        IF (CartesianVx > VXThreshold)
           AND (CartesianForcefX > FXThreshold) THEN

            CASE stFromUnity.nGameStatus OF

                0: // Not playing
                    stJointTargetTorque.M1 := 0.0;

                1: // Light bin
                    stJointTargetTorque.M1 := 0.0;

                2: // Medium bin
                    stJointTargetTorque.M1 := 7.0;

                3: // Heavy bin
                    stJointTargetTorque.M1 := 15.0;

                ELSE
                    stJointTargetTorque.M1 := 0.0;

            END_CASE;


        (****************************************************
            CONDITION 2: NEGATIVE X MOVEMENT

            Both Vx and Fx must be negative
            and below their negative thresholds.

            Apply POSITIVE resistance.
        *****************************************************)

        ELSIF (CartesianVx < -VXThreshold)
              AND (CartesianForcefX < -FXThreshold) THEN

            CASE stFromUnity.nGameStatus OF

                0: // Not playing
                    stJointTargetTorque.M1 := 0.0;

                1: // Light bin
                    stJointTargetTorque.M1 := 0.0;

                2: // Medium bin
                    stJointTargetTorque.M1 := -7.0;

                3: // Heavy bin
                    stJointTargetTorque.M1 := -15.0;

                ELSE
                    stJointTargetTorque.M1 := 0.0;

            END_CASE;

        ELSE

            // Force and velocity conditions not satisfied
            stJointTargetTorque.M1 := 0.0;

        END_IF;
	
	ELSE
		
		GVL_HMI.bLaunchGameSorter:= FALSE;
	
	END_IF

  

END_IF;

END_FUNCTION_BLOCK

// ---- POUs/Crazy Car/FB_CrazyCarGame.TcPOU
FUNCTION_BLOCK FB_CrazyCarGame

VAR_INPUT
    bEnable                   : BOOL;
    stCartesianPosePercentage : ST_CartesianPose;
    fWristAngleDeg            : LREAL;
    CartesianVtheta           : LREAL;
    CartesianMtheta           : LREAL;
END_VAR

VAR_OUTPUT
    stJointTargetTorque : ST_JointTorque;
END_VAR

VAR
    // =====================================================
    // UNITY COMMUNICATION
    // =====================================================

    stToUnity   : ST_CrazyCarToUnity;
    stFromUnity : ST_UnityToCrazyCar;


    // =====================================================
    // RESISTANCE LEVELS
    // =====================================================

    TorqueTaxi  : LREAL := 0.0;
    TorqueVan   : LREAL := 20.0;
    TorqueTruck : LREAL := 40.0;

    TorqueSign  : LREAL := 1.0;

    fTorque : LREAL := 0.0;


    // =====================================================
    // VELOCITY FILTER
    // =====================================================

    fVthetaFiltered : LREAL := 0.0;

    fFilterTime : LREAL := 0.015;

    fTaskCycleTime : LREAL := 0.01;


    // =====================================================
    // VELOCITY DEAD ZONE AND TRANSITION
    //
    // Assumes CartesianVtheta is in deg/s
    // =====================================================

    fVelocityDeadband : LREAL := 10.0;

    fVelocityFull : LREAL := 30.0;


    // =====================================================
    // SMOOTH RESISTANCE
    // =====================================================

    fVelocityMagnitude : LREAL := 0.0;

    fVelocityFactor : LREAL := 0.0;

    fSmoothFactor : LREAL := 0.0;

    fTorqueTarget : LREAL := 0.0;

    fTorqueCommand : LREAL := 0.0;


    // =====================================================
    // APPLICATION TORQUE SLEW LIMIT
    //
    // Units must match the game torque command per second.
    // =====================================================

    fTorqueRateLimit : LREAL := 100.0;

    fMaxTorqueStep : LREAL := 0.0;

    fTorqueDifference : LREAL := 0.0;


    // =====================================================
    // INITIAL BENCH-TEST LIMITS
    //
    // Keep motor output disabled while validating the logic.
    // fMaxGameTorque is an experimental command bound,
    // NOT a validated safe human-interaction torque.
    // =====================================================

    bEnableResistanceOutput : BOOL := FALSE;

    fMaxGameTorque : LREAL :=40.0;

END_VAR

(************************************************************
    CRAZY CAR GAME - CONTINUOUS SMOOTH RESISTANCE

    Unity status:
        0 = Menu / Popup
        1 = Taxi
        2 = Van
        3 = Truck

    Objectives:
        1. Zero resistance near stationary velocity
        2. Smooth resistance transition
        3. Approximately constant resistance during motion
        4. Avoid binary torque switching
        5. Limit the commanded torque rate
*************************************************************)


// ==========================================================
// 1. DEFAULT OUTPUTS
// ==========================================================

stJointTargetTorque.M1 := 0.0;
stJointTargetTorque.M2 := 0.0;
stJointTargetTorque.M3 := 0.0;

stToUnity.GameIsActive := FALSE;

fTorque := 0.0;
fTorqueTarget := 0.0;


// ==========================================================
// 2. CHECK GAME ENABLE
// ==========================================================

IF bEnable AND NOT stFromUnity.bGameClosed THEN

    // Send data to Unity

    stToUnity.fY :=
        LREAL_TO_REAL(stCartesianPosePercentage.Y);

    stToUnity.fWristAngle :=
        LREAL_TO_REAL(fWristAngleDeg);

    stToUnity.GameIsActive := TRUE;


    // ======================================================
    // 3. READ VEHICLE RESISTANCE
    // ======================================================

    CASE stFromUnity.nGameStatus OF

        1:
            fTorque := TorqueTaxi;

        2:
            fTorque := TorqueVan;

        3:
            fTorque := TorqueTruck;

        ELSE
            fTorque := 0.0;

    END_CASE;


    // ======================================================
    // 4. FILTER WRIST VELOCITY
    // ======================================================

    IF (fTaskCycleTime > 0.0)
       AND (fFilterTime >= 0.0) THEN

        fVthetaFiltered :=
            fVthetaFiltered
            +
            (
                fTaskCycleTime /
                (fFilterTime + fTaskCycleTime)
            )
            *
            (CartesianVtheta - fVthetaFiltered);

    ELSE

        fVthetaFiltered := 0.0;

    END_IF;


    // ======================================================
    // 5. CALCULATE VELOCITY MAGNITUDE
    // ======================================================

    fVelocityMagnitude := ABS(fVthetaFiltered);


    // ======================================================
    // 6. CALCULATE CONTINUOUS VELOCITY FACTOR
    //
    // Dead zone:          Factor = 0
    // Transition region:  Factor = 0..1
    // Full movement:      Factor = 1
    // ======================================================

    fVelocityFactor := 0.0;

    IF fVelocityFull > fVelocityDeadband THEN

        IF fVelocityMagnitude <= fVelocityDeadband THEN

            fVelocityFactor := 0.0;

        ELSIF fVelocityMagnitude >= fVelocityFull THEN

            fVelocityFactor := 1.0;

        ELSE

            fVelocityFactor :=
                (fVelocityMagnitude - fVelocityDeadband)
                /
                (fVelocityFull - fVelocityDeadband);

        END_IF;

    END_IF;


    // ======================================================
    // 7. SMOOTHSTEP FUNCTION
    //
    // Smooth transition from 0 to 1.
    //
    // f(x) = 3*x*x - 2*x*x*x
    //
    // This avoids an abrupt slope change at the
    // beginning and end of the transition region.
    // ======================================================

    fSmoothFactor :=
        fVelocityFactor
        *
        fVelocityFactor
        *
        (3.0 - 2.0 * fVelocityFactor);


    // ======================================================
    // 8. CALCULATE TARGET RESISTANCE
    //
    // Preserve your existing motor sign convention.
    // Verify that the physical wrist torque opposes motion.
    // ======================================================

    IF fVthetaFiltered > fVelocityDeadband THEN

        fTorqueTarget :=
            TorqueSign
            *
            fTorque
            *
            fSmoothFactor;

    ELSIF fVthetaFiltered < -fVelocityDeadband THEN

        fTorqueTarget :=
            -TorqueSign
            *
            fTorque
            *
            fSmoothFactor;

    ELSE

        fTorqueTarget := 0.0;

    END_IF;


    // ======================================================
    // 9. LIMIT GAME TORQUE MAGNITUDE
    //
    // Experimental bench-test limit.
    // ======================================================

    IF bEnableResistanceOutput
       AND (fMaxGameTorque > 0.0) THEN

        fTorqueTarget :=
            MAX(
                -fMaxGameTorque,
                MIN(fMaxGameTorque, fTorqueTarget)
            );

    ELSE

        fTorqueTarget := 0.0;

    END_IF;


    // ======================================================
    // 10. APPLICATION-LEVEL TORQUE SLEW LIMIT
    //
    // Prevent large command changes within one PLC cycle.
    // ======================================================

    fMaxTorqueStep :=
        MAX(0.0, fTorqueRateLimit)
        *
        MAX(0.0, fTaskCycleTime);

    fTorqueDifference :=
        fTorqueTarget - fTorqueCommand;


    IF fTorqueDifference > fMaxTorqueStep THEN

        fTorqueCommand :=
            fTorqueCommand + fMaxTorqueStep;

    ELSIF fTorqueDifference < -fMaxTorqueStep THEN

        fTorqueCommand :=
            fTorqueCommand - fMaxTorqueStep;

    ELSE

        fTorqueCommand := fTorqueTarget;

    END_IF;


    // ======================================================
    // 11. TRANSFER TORQUE TO WRIST MOTORS
    // ======================================================

    IF bEnableResistanceOutput THEN

        stJointTargetTorque.M2 := fTorqueCommand;
        stJointTargetTorque.M3 := fTorqueCommand;

    ELSE

        stJointTargetTorque.M2 := 0.0;
        stJointTargetTorque.M3 := 0.0;

        fTorqueCommand := 0.0;

    END_IF;


ELSE

    // ======================================================
    // 12. GAME DISABLED OR CLOSED
    // ======================================================

    IF bEnable AND stFromUnity.bGameClosed THEN

        GVL_HMI.bLaunchGameCrazyCar := FALSE;

    END_IF;


    stToUnity.GameIsActive := FALSE;

    fTorque := 0.0;
    fTorqueTarget := 0.0;
    fTorqueCommand := 0.0;

    fVthetaFiltered := 0.0;

    fVelocityMagnitude := 0.0;
    fVelocityFactor := 0.0;
    fSmoothFactor := 0.0;

    fTorqueDifference := 0.0;

END_IF;

END_FUNCTION_BLOCK

// ---- POUs/Firrfly Game/FB_FireflyGame.TcPOU
FUNCTION_BLOCK FB_FireflyGame
VAR_INPUT
    bEnable                   : BOOL;
    stCartesianPosePercentage : ST_CartesianPose; // from Kinematics: X -100..+100 %, Y 0..100 % (0..370 mm)
END_VAR
VAR_OUTPUT
    stJointTargetTorque : ST_JointTorque;  // always 0: Firefly is motion-only, no actuation
    nGameStatus         : INT;             // Unity game status, for MAIN / HMI
    bExitRequested      : BOOL;            // TRUE for ONE PLC cycle when Exit is pressed in Unity
    bWrongFlowerEvent   : BOOL;            // TRUE for ONE PLC cycle per wrong flower (for later haptics)
END_VAR
VAR
    stToUnity   : ST_FireflyToUnity;
    stFromUnity : ST_FireflyFromUnity;

    // Calibration: robot percent (from Kinematics) at home, and travel either side of home
    // that brings the firefly to the edge of the garden (= +/-100 % in Unity).
    fXHome      : REAL := 0.0;    // X percent at home (middle of the workspace)
    fYHome      : REAL := 50.0;   // Y percent at home (middle of 0..370 mm = 185 mm)
    fXHalfRange : REAL := 50.0;   // X: lower this if X needs less motion than Y
    fYHalfRange : REAL := 25.0;   // Y: +/-25 % = 50 % of the Y range of motion in total

    rtExit  : R_TRIG;
    rtWrong : R_TRIG;
    fXRaw   : REAL;
    fYRaw   : REAL;
END_VAR

// Firefly is motion-only: never apply torque.
stJointTargetTorque.M1 := 0.0;
stJointTargetTorque.M2 := 0.0;
stJointTargetTorque.M3 := 0.0;

IF bEnable THEN
    fXRaw := TO_REAL(stCartesianPosePercentage.X);
    fYRaw := TO_REAL(stCartesianPosePercentage.Y);
    // Home -> 0 %, home +/- half range -> +/-100 %, clamped so the firefly stays inside the garden.
    stToUnity.fX := LIMIT(-100.0, (fXRaw - fXHome) / MAX(fXHalfRange, 0.1) * 100.0, 100.0);
    stToUnity.fY := LIMIT(-100.0, (fYRaw - fYHome) / MAX(fYHalfRange, 0.1) * 100.0, 100.0);
ELSE
    stToUnity.fX := 0.0;   // firefly waits on the home flower
    stToUnity.fY := 0.0;
END_IF

// Unity's pulses -> one-cycle events for MAIN (each new pulse = a new rising edge).
rtExit(CLK := stFromUnity.bExitPressed);
rtWrong(CLK := stFromUnity.bWrongFlower);
bExitRequested    := rtExit.Q;
bWrongFlowerEvent := rtWrong.Q;
nGameStatus       := stFromUnity.nGameStatus;

END_FUNCTION_BLOCK

// ---- POUs/FB_ForceTorqueSensor.TcPOU
FUNCTION_BLOCK FB_ForceTorqueSensor
VAR_IN_OUT
 CartesianState : ST_CartesianState;
 
END_VAR
VAR_INPUT
	CartesianPosAdditionalParameter :ST_CartesianAdditionalParametes;
END_VAR
VAR
    eState : E_CalibrationState :=  E_CalibrationState.INIT;
    tWait  : TON;
	FxTemp : LREAL;
	FyTemp : LREAL;
	MzTemp : LREAL;
	OffsetRawFx: LINT;
	OffsetRawFy: LINT;
	OffsetRawMz: LINT;
	sumFx: LINT;
	sumFy: LINT;
	sumMz: LINT;
	nSample: INT;
	rTrigZero : R_TRIG;
	Theta1: LREAL;
	Theta2: LREAL;
	Theta3: LREAL;
END_VAR
VAR CONSTANT
    CMD_STOP   : DWORD := 16#0000000C;
    CMD_FILTER : DWORD := 16#00050108;  // 1st-order LPF, 100 Hz
    CMD_START  : DWORD := 16#0000000B;
    FORCE_DIV  : REAL := 50.0;     // RFT60-HA01 force divider
	TORQUE_DIV : REAL := 2000.0;   // RFT60-HA01 torque divider
	CostanstAngleBetweenFTSensorAndXdirection : LREAL := 30.0; // Unit Degree
	CostanstAngleBetweenFTSensorAndYdirection : LREAL := 30.0; // Unit Degree
	ZeroingSample : INT := 100;
	
END_VAR



CASE eState OF
E_CalibrationState.INIT:
    GVL_ForceTorqueSensor.ConfigParameter := CMD_STOP;
    tWait(IN := TRUE, PT := T#1000MS);
    IF tWait.Q THEN tWait(IN := FALSE); eState := E_CalibrationState.SET_FILTER; END_IF

E_CalibrationState.SET_FILTER:
   GVL_ForceTorqueSensor.ConfigParameter := CMD_FILTER;
    tWait(IN := TRUE, PT := T#1000MS);
    IF tWait.Q THEN tWait(IN := FALSE); eState := E_CalibrationState.START; END_IF

E_CalibrationState.START:
    GVL_ForceTorqueSensor.ConfigParameter := CMD_START;
    eState := E_CalibrationState.WaitingforCalibrationButton;
	sumFx := 0; sumFy := 0;  sumMz := 0;
	
E_CalibrationState.WaitingforCalibrationButton:

rTrigZero(CLK := GVL_HMI.StartCalibrationButton);

IF rTrigZero.Q THEN

    
   
    GVL_HMI.StartCalibrationButton := FALSE;
	eState := E_CalibrationState.ZEROING;
	sumFx := 0;
	sumFy := 0;
	sumMz := 0;
	nSample := 0;
	tWait(IN := FALSE);   // reset timer

END_IF

	
E_CalibrationState.ZEROING:
   

	tWait(IN := TRUE, PT := T#2000MS);          // let streaming/filter settle first
    IF tWait.Q THEN
        sumFx := sumFx + GVL_ForceTorqueSensor.RawFx;
        sumFy := sumFy + GVL_ForceTorqueSensor.RawFy;
        sumMz := sumMz + GVL_ForceTorqueSensor.RawMz;
        nSample := nSample + 1;
        IF nSample >= ZeroingSample THEN
            OffsetRawFx := sumFx / ZeroingSample;
            OffsetRawFy := sumFy / ZeroingSample;
            OffsetRawMz := sumMz / ZeroingSample;
            eState := E_CalibrationState.RUNNING;
        END_IF
    END_IF



E_CalibrationState.RUNNING:
IF GVL_HMI.StartCalibrationButton THEN
	 GVL_HMI.StartCalibrationButton := FALSE;

    sumFx := 0;
    sumFy := 0;
    sumMz := 0;
    nSample := 0;

    tWait(IN := FALSE);

    eState := E_CalibrationState.ZEROING;
END_IF
// All Angles that is used for rotational frames;
Theta1:= CostanstAngleBetweenFTSensorAndXdirection;   //UNIT: degree   Shift for F/t Sensor, it is related to design and I got from SOLIDWORKS// this number is constant;
Theta2 := -CartesianPosAdditionalParameter.BetaIncremental; // UNIT: degree  the angle between frame x,y with refrence
Theta3 := -Cartesianstate.Position.Theta; //UNIT: degree  the wrist angle between x-frame of wrist with x-frame of reference
//
    FxTemp := LINT_TO_REAL(GVL_ForceTorqueSensor.RawFx- OffsetRawFx) / FORCE_DIV;
    FyTemp := LINT_TO_REAL(GVL_ForceTorqueSensor.RawFy-OffsetRawFy) / FORCE_DIV;
    MzTemp := LINT_TO_REAL(GVL_ForceTorqueSensor.RawMz-OffsetRawMz) / TORQUE_DIV;
	CartesianState.Force.Fx :=-( FxTemp * COS((Theta1 + Theta2 + Theta3)*(PI / 180.0))-
	FyTemp * SIN((Theta1 + Theta2 + Theta3)*(PI / 180.0)));
	
	GVL_HMI.Fx_HMI := CartesianState.Force.Fx ; // Display in HMI
	
	CartesianState.Force.Fy := -(FxTemp * SIN((Theta1 + Theta2 + Theta3)*(PI / 180.0))+
	FyTemp * COS((Theta1 + Theta2 + Theta3)*(PI / 180.0)));
	
	GVL_HMI.Fy_HMI := CartesianState.Force.Fy; // Display in HMI
	CartesianState.Force.Mtheta := MzTemp ;
	GVL_HMI.Mz_HMI := CartesianState.Force.Mtheta*1000;  // Display in HMI //Unit : mNM




END_CASE

IF eState = E_CalibrationState.RUNNING THEN
	GVL_HMI.UserSecuringButton_HMI := TRUE;
	ELSE
	GVL_HMI.UserSecuringButton_HMI := FALSE;	
END_IF

END_FUNCTION_BLOCK

// ---- POUs/HMI_FunBlock/MicroswitchCheck.TcPOU
FUNCTION_BLOCK MicroswitchCheck
VAR_INPUT
END_VAR
VAR_OUTPUT
END_VAR
VAR
	SwTheta1: BOOL;
	SwTheta2: BOOL;
	SwR1: BOOL;
	SwR2: BOOL;
	SwBeta1: BOOL;
	SwBeta2: BOOL;
END_VAR

SwTheta1 	 := (GVL_MicroSwitch.dwMicroSwitchDriverA AND 16#00020000) <> 0;  (* bit 0 *)
SwTheta2     := (GVL_MicroSwitch.dwMicroSwitchDriverA AND 16#00010000) <> 0;  (* bit 1 *)
SwR1    	 := (GVL_MicroSwitch.dwMicroSwitchDriverB AND 16#00080000) <> 0;  (* bit 0 *)
SwR2  		 := (GVL_MicroSwitch.dwMicroSwitchDriverB AND 16#00040000) <> 0;  (* bit 1 *)
SwBeta1      := (GVL_MicroSwitch.dwMicroSwitchDriverB AND 16#00020000) <> 0;  (* bit 2 *)
SwBeta2      := (GVL_MicroSwitch.dwMicroSwitchDriverB AND 16#00010000) <> 0;  (* bit 3 *)

IF SwTheta1 THEN
GVL_HMI.CheckMicroswitchWristLeft := TRUE;
	
END_IF

IF SwTheta2 THEN
GVL_HMI.CheckMicroswitchWristRight := TRUE;
	
END_IF

IF SwR1 THEN
GVL_HMI.CheckMicroswitchLinearMax := TRUE;
	
END_IF

IF SwR2 THEN
GVL_HMI.CheckMicroswitchLinearMin := TRUE;
	
END_IF

IF SwBeta1 THEN
GVL_HMI.CheckMicroswitchRotationRight := TRUE;
	
END_IF

IF SwBeta2 THEN
GVL_HMI.CheckMicroswitchRotationLeft := TRUE;
	
END_IF

IF GVL_HMI.CheckMicroswitchWristLeft AND GVL_HMI.CheckMicroswitchWristRight AND GVL_HMI.CheckMicroswitchLinearMax AND GVL_HMI.CheckMicroswitchLinearMin AND GVL_HMI.CheckMicroswitchRotationRight AND GVL_HMI.CheckMicroswitchRotationLeft THEN
GVL_HMI.ContinueToHoming := TRUE;

END_IF

END_FUNCTION_BLOCK

// ---- POUs/HMI_FunBlock/FB_UserSecuring.TcPOU
FUNCTION_BLOCK FB_UserSecuring
VAR_INPUT
END_VAR
VAR_OUTPUT
END_VAR
VAR
END_VAR

IF GVL_HMI.check1 AND GVL_HMI.check2 AND GVL_HMI.check3 AND GVL_HMI.check4 AND GVL_HMI.check5 AND GVL_HMI.check6 THEN
	
GVL_HMI.ContinueTOWorkspaceLimits := TRUE;
ELSE
	
GVL_HMI.ContinueTOWorkspaceLimits := FALSE;

END_IF

END_FUNCTION_BLOCK

// ---- POUs/FB_TherapyManager.TcPOU
FUNCTION_BLOCK FB_TherapyManager

VAR_INPUT
	Enable         : BOOL;
    Config         : ST_TherapyConfig;       // The struct we just built!
    ActualJoints    : ST_JointState;        // Feedback: Joint q, q_dot, M
    ActualCartesian : ST_CartesianState;    // Feedback: Cartesian Pose, Vel, Force
    TargetCartesian : ST_CartesianTarget;   // Target: Cartesian Pose, Vel, Force setpoints
    SimpleJointTorqueObtainedFromGames : ST_JointTorque;
    fbKinematics    : REFERENCE TO FB_RobotKinematics;
	WallSetPointXandY : ARRAY[1..4, 1..2] OF LREAL;
END_VAR
VAR_OUTPUT
	TargetJointsTorque    : ST_JointTorque;        // Output for CST Mode
	//TargetMode      : En_TargetMode;              // Drive mode (eCSP, eCSV, eCST)
    //  Out_Positions  : ST_JointPositions;      // Output for CSV Mode
END_VAR
VAR
	// 1. The Expert Math Blocks
    fbImpedance    : FB_ImpedanceController;
    fbAdmittance   : FB_AdmittanceController;
	fbForceYield : FB_ForceController;
    fbDynamics     : FB_DynamicsCompensator;
    
    // 2. Internal Routing Variables
    TherapyForces   : ST_CartesianForces;             // Cartesian Space (End-Effector force)
    TherapyTorque   : ST_JointTorque;                 // Joint Space (Therapy motor torque)
    CompTorque      : ST_JointTorque;                 // Joint Space (Hardware compensation torque)
	timerHold : TON;
	
	// Wall Variables
	WallTorque : ST_JointTorque;
	fbVirtualWall : FB_VirtuallWall;
	bWallInContact : BOOL;
	WallCartesianForce: ST_CartesianForces;
	MotionState: INT := 1;
	//cycle: INT;
	CycleMotion: INT :=1;
	
	
	fbMicroswitchCheck : MicroswitchCheck;   // Delete this after cycling test
	fbStopM1 : MC_Stop;
	fbStopM2 : MC_Stop;
	fbStopM3 : MC_Stop;
	firsttime: BOOL := TRUE;
END_VAR
VAR CONSTANT
    // Zero constants for clean single-line memory resets
    cZeroTorque : ST_JointTorque    := (M1 := 0.0, M2 := 0.0, M3 := 0.0);
    cZeroForces : ST_CartesianForces := (Fx := 0.0, Fy := 0.0, Mtheta := 0.0);
END_VAR

// =========================================================
// 1. SAFETY DISABLE GUARD
// =========================================================
IF NOT Enable THEN
    TargetJointsTorque := cZeroTorque;
	
   
    RETURN;
END_IF

// =========================================================
// 2. CLEAR INTERMEDIATE BUFFERS (PREVENT STALE DATA LEAKS)
// =========================================================
TherapyForces := cZeroForces;
TherapyTorque := cZeroTorque;
WallTorque := cZeroTorque;
CompTorque    := cZeroTorque;

// =========================================================
// 3. PRIMARY CONTROLLER ROUTING
// =========================================================
CASE Config.ControllerType OF

    E_ControllerType.ControlNone:
        TherapyTorque := SimpleJointTorqueObtainedFromGames;
		
		(*

    E_ControllerType.ControlImpedance:
        // Step A: Virtual spring-damper computes interaction forces
        fbImpedance(
            Stiffness   := Config.Stiffness_K,
            Damping     := Config.Damping_D,
            ActualPose  := ActualCartesian.Position,
            TargetPose  := TargetCartesian.Position,
            ActualVel   := ActualCartesian.Velocity,
            TargetVel   := TargetCartesian.Velocity,
            OutputForce => TherapyForces
        );
        
        // Step B: Map Cartesian Force -> Joint Torque via J^T
        TherapyTorque := fbKinematics.ApplyJacobianTranspose(Force := TherapyForces);

    E_ControllerType.ControlAdmittance:
        // Measured patient forces generate target positions / velocities
        fbAdmittance(
            TherapyMode     := Config.TherapyMode,
            VirtualMass     := Config.Mass_M,
            VirtualDamp     := Config.Damping_D,
            MeasuredForces  := ActualCartesian.Forces,
            TargetForces    := TargetCartesian.Forces,
            ActualPose      := ActualCartesian.Position,
            TargetPosition  => TargetJoints.Position
        );

    E_ControllerType.ControlForce:
        // Generic Yield-Threshold / Breakaway Force Controller
        fbForceYield(
            ForceThreshold := Config.ForceConfig.Threshold, // Generic resistance force
            VirtualDamping := Config.ForceConfig.Damping,   // Generic motion viscosity
            ActualForce    := ActualCartesian.Forces,
            ActualJoints   := ActualJoints,
            OutputTorque   => TherapyTorque
        );
		*)

END_CASE

// =========================================================
// 4. HARDWARE DYNAMICS COMPENSATION (Joint Space)
// =========================================================

(*

IF Config.FeatureFrictionComp OR Config.FeatureInertiaComp OR Config.FeatureGravityComp THEN
    fbDynamics(
        JointPosition  := ActualJoints.Position,
        JointVelocity  := ActualJoints.Velocity,
        EnableGravity  := Config.FeatureGravityComp,
        EnableFriction := Config.FeatureFrictionComp,
        EnableInertia  := Config.FeatureInertiaComp,
        CompTorque     => CompTorque
    );
END_IF
*)
// Cycle Test
(* 

IF  firsttime THEN
GVL_hmi.CheckMicroswitchLinearMax := FALSE;
GVL_hmi.CheckMicroswitchLinearMin := FALSE;
GVL_hmi.CheckMicroswitchRotationLeft := FALSE;
GVL_hmi.CheckMicroswitchRotationRight := FALSE;
GVL_HMI.CheckMicroswitchWristLeft := FALSE;
GVL_HMI.CheckMicroswitchWristRight := FALSE;
firsttime := FALSE;
END_IF
// Tests
fbMicroswitchCheck();
IF GVL_hmi.CheckMicroswitchLinearMax OR GVL_hmi.CheckMicroswitchLinearMin OR
 GVL_hmi.CheckMicroswitchRotationLeft OR GVL_hmi.CheckMicroswitchRotationRight OR 
 GVL_HMI.CheckMicroswitchWristLeft OR GVL_HMI.CheckMicroswitchWristRight

THEN
 
	fbStopM1(
        Axis      := GVL_Axes.Axis1,
        Execute   := TRUE);   

    fbStopM2(
        Axis      := GVL_Axes.Axis2,
        Execute   := TRUE);

    fbStopM3(
        Axis      := GVL_Axes.Axis3,
        Execute   := TRUE);
END_IF

CASE MotionState OF
	1: // Motor1 +_
		TherapyTorque.M1 := -8.0;
		TherapyTorque.M2 := 0.0;
		TherapyTorque.M3 := 0.0;
		IF ActualCartesian.Position.X> 200.0 THEN
			
		TherapyTorque.M1 :=  0.05* ActualCartesian.Velocity.Vx;
		TherapyTorque.M2 := 0.0;
		TherapyTorque.M3 := 0.0;
		timerHold(IN := TRUE, PT := T#1S);
		
		IF timerHold.Q THEN
            timerHold(IN := FALSE); // Reset the timer so it can be reused later
            MotionState := 2;
        END_IF
			
		END_IF
	2: // linear +
		TherapyTorque.M1 := 0.0;
		TherapyTorque.M2 := 8.0;
		TherapyTorque.M3 := -8.0;
		
		IF ActualCartesian.Position.Y> 300.0 THEN
		TherapyTorque.M1 := 0.0;
		TherapyTorque.M2 :=  - 0.05* ActualCartesian.Velocity.Vy;
		TherapyTorque.M3 :=  0.05* ActualCartesian.Velocity.Vy;
		timerHold(IN := TRUE, PT := T#1S);
		
		IF timerHold.Q THEN
            timerHold(IN := FALSE); // Reset the timer so it can be reused later
            MotionState := 3;
		END_IF
		END_IF
	 3: // Motor1 -
		TherapyTorque.M1 := 8.0;
		TherapyTorque.M2 := 0.0;
		TherapyTorque.M3 := 0.0;
		
		IF ActualCartesian.Position.X< -50.0 THEN
		TherapyTorque.M1 := 0.05* ActualCartesian.Velocity.Vx;
		TherapyTorque.M2:= 0.0;
		TherapyTorque.M3 := 0.0;
		timerHold(IN := TRUE, PT := T#1S);
		
		IF timerHold.Q THEN
            timerHold(IN := FALSE); // Reset the timer so it can be reused later
            MotionState := 4;
		END_IF
		END_IF
	 4: // linear -
		TherapyTorque.M1 := 0.0;
		TherapyTorque.M2 := -8.0;
		TherapyTorque.M3 := 8.0;
		
		
		IF ActualCartesian.Position.Y< 150.0 THEN
		TherapyTorque.M1 := 0.0;
		TherapyTorque.M2 :=  - 0.05* ActualCartesian.Velocity.Vy;
		TherapyTorque.M3 :=  0.05* ActualCartesian.Velocity.Vy;
		timerHold(IN := TRUE, PT := T#1S);
		
		IF timerHold.Q THEN
            timerHold(IN := FALSE); // Reset the timer so it can be reused later
			CycleMotion := CycleMotion+1;
		IF CycleMotion = 500 THEN
            MotionState := 5;
		ELSE
	MotionState := 1;
			
		END_IF
		END_IF
		END_IF
		
		
	 5: 
		TherapyTorque.M1 := 0.0;
		TherapyTorque.M2 := 0.0;
		TherapyTorque.M3 := 0.0;
		
	 
	 
	
END_CASE

*)// Cycle Test

// VirtualWallTorque

fbVirtualWall(
    bEnable     := GVL_HMI.EableVirtuallWall_Planar,
	Endeffectorstatus := ActualCartesian,
	WallSetPointXandY := WallSetPointXandY,
	WallCartesianForce => WallCartesianForce,
	bInContact  => bWallInContact
    
);

WallTorque :=
    fbKinematics.CartesianForceToTorque(
        Force := WallCartesianForce
    );





// =========================================================
// 5. FINAL TORQUE SUMMATION & GLOBAL SAFETY CLAMP
// =========================================================
IF bWallInContact THEN

    // Virtual wall is active:
    // use wall torque only
    TargetJointsTorque.M1 := LIMIT(
        -Config.GlobalForceLimit,
        WallTorque.M1,
        Config.GlobalForceLimit
    );

    TargetJointsTorque.M2 := LIMIT(
        -Config.GlobalForceLimit,
        WallTorque.M2,
        Config.GlobalForceLimit
    );

    TargetJointsTorque.M3 := LIMIT(
        -Config.GlobalForceLimit,
        WallTorque.M3,
        Config.GlobalForceLimit
    );

ELSE

    // No wall contact:
    // normal robot torque
    TargetJointsTorque.M1 := LIMIT(
        -Config.GlobalForceLimit,
        TherapyTorque.M1 + CompTorque.M1,
        Config.GlobalForceLimit
    );

    TargetJointsTorque.M2 := LIMIT(
        -Config.GlobalForceLimit,
        TherapyTorque.M2 + CompTorque.M2,
        Config.GlobalForceLimit
    );

    TargetJointsTorque.M3 := LIMIT(
        -Config.GlobalForceLimit,
        TherapyTorque.M3 + CompTorque.M3,
        Config.GlobalForceLimit
    );

END_IF;

END_FUNCTION_BLOCK

// ---- POUs/FB_ImpedanceController.TcPOU
FUNCTION_BLOCK FB_ImpedanceController
VAR_INPUT
 TherapyMode : E_RehabMode;
 Stiffness   : LREAL;              // Virtual spring K
 Damping     : LREAL;              // Virtual friction D
  
END_VAR



VAR_OUTPUT
    bBusy         : BOOL;
    bError        : BOOL;
    bDone         : BOOL;
//	TherapyTorques : ST_JointTorques;
END_VAR

VAR
	 
    stPointA      : ARRAY [1..3] OF LREAL  ; 
    stPointB      : ARRAY [1..3] OF LREAL  ;
    stPointC      : ARRAY [1..3] OF LREAL  ;
	
    // --- Feedback from Robot (Inputs) ---
    ActX          : LREAL; 
    ActY          : LREAL; 
    ActTheta      : LREAL;
	ActR          : LREAL; // mm
	ActBeta		  : LREAL;
    


    // --- State Machine Logic ---
    iState           : INT := 0;      // Main Step Counter
    iCurrentSegment  : INT := 0;      // 5=Approach, 10=A->B, 20=B->C, 30=C->A
    bAtPointA        : BOOL := FALSE;
    bSegmentDone     : BOOL;
    bWaitEnable      : BOOL;
    
    // --- Timers & Sub-FBs ---
    fbWaitTimer      : TON;           // Timer for resting at corners
    fbKinematic      : FB_RobotKinematics;  // Internal instance to update kinematics
    
    // --- Motion Profile Variables (Trapezoid Generator) ---
    lrS_T            : LREAL;         // Current Distance along path (0 to L)
    lrS_dot          : LREAL;         // Current Velocity (Speed of the "Rabbit")
    lrL_Target       : LREAL;         // Total Length of the current segment

    // --- Geometric Calculations (Approach Phase) ---
    lrApproachStartX : LREAL;
    lrApproachStartY : LREAL;
    lrApproachStartTheta : LREAL;
    lrDX_App, lrDY_App, lrDTh_App, lrL_App : LREAL;

    // --- Geometric Calculations (Triangle Phase) ---
    // Line 1 (A->B)
    lrDX1, lrDY1, lrDTh1, lrL1 : LREAL;
    // Line 2 (B->C)
    lrDX2, lrDY2, lrDTh2, lrL2 : LREAL;
    // Line 3 (C->A)
    lrDX3, lrDY3, lrDTh3, lrL3 : LREAL;

    // --- Impedance Control Targets ---
    SetAppX             : LREAL; // The "Virtual Rabbit" X position
    SetAppY             : LREAL; // The "Virtual Rabbit" Y position
    SetAppTheta         : LREAL; // The "Virtual Rabbit" Theta position
    
    // --- Calculation Results ---
    CalcForces       : ARRAY [1..3] OF LREAL; // [Fx, Fy, Mz] calculated by Impedance
    CalcTorques      : ARRAY [1..3] OF LREAL; // [Tau1, Tau2, Tau3] calculated by Jacobian

    // --- TwinCAT Motion Control Blocks ---
    // Note: I renamed these to 'fbTorqueAxis1' to match the method code we wrote previously
    fbTorqueAxis1    : MC_TorqueControl;
    fbTorqueAxis2    : MC_TorqueControl;
    fbTorqueAxis3    : MC_TorqueControl;

    // --- Safety Parameters ---
    MaxSpeedLimit    : LREAL := 70.0; // Safety velocity limit (mm/s)
    MaxTorqueLimit   : LREAL := 50.0;  // Safety torque limit (Nm)
	
	// 
	lrVmax: LREAL := 10.0; // mm/s
	lrAcc : LREAL := 100.0 ;// mm/ s^2
	
	SetVelAppX      : LREAL;
    SetVelAppY      : LREAL;
    SetVelAppTheta  : LREAL;
	
	// INTERNAL setpoints calculated each cycle
    stCurrentSet  : ARRAY[1..3] OF LREAL; // Target [X, Y, Theta]
	 lrVx_FF, lrVy_FF, lrVTh_FF : LREAL;
	  Ex, Ey, ETheta    : LREAL; // Position Errors
	  lrTorqueSetpoint_Pct : ARRAY[1..3] OF LREAL;
END_VAR

(* This Function block can be used for difference rehabilitation mode
 1- passive motion: actuators create No torque and patient can move the robot
 2- Passive motion + Compensation(solving dynamic of robot)
 3- Resistive or Assistive force
*)

stPointA := GVL_TargetPoints.Target_A;
stPointB := GVL_TargetPoints.Target_B;
stPointC := GVL_TargetPoints.Target_C;


// =========================================================
// 1. KINEMATICS UPDATE (Always Run First)
// =========================================================
// We need ActX/ActY to calculate the spring force error
(*  JUST FOR TEST ELIMINATED
fbKinematic(
	
    q1 := GVL_RobotData.Q1_Actual, 
    q2 := GVL_RobotData.Q2_Actual, 
    q3 := GVL_RobotData.Q3_Actual, 
    X_Dir => ActX, 
    Y_Dir => ActY, 
    Theta => ActTheta,
    R_Dir => ActR,
	Beta => ActBeta    
);
*)

// 

// Update Timer
fbWaitTimer(IN := bWaitEnable, PT := T#120S);

// =========================================================
// 2. STATE MACHINE
// =========================================================
CASE iState OF

    // -----------------------------------------------------
    // STATE 0: INITIALIZATION (Math Setup)
    // -----------------------------------------------------
    0: 
        // 1. Capture Start Position for Approach
        lrApproachStartX     := ActX;
        lrApproachStartY     := ActY;
        lrApproachStartTheta := ActTheta;

        // 2. Calculate Distance to Point A (Approach Vector)
        lrDX_App  := stPointA[1] - lrApproachStartX;
        lrDY_App  := stPointA[2] - lrApproachStartY;
        lrDTh_App := stPointA[3] - lrApproachStartTheta;
        lrL_App   := MAX(0.001, SQRT(lrDX_App*lrDX_App + lrDY_App*lrDY_App));

        // 3. Calculate Triangle Vectors (A->B, B->C, C->A)
        // --- Line 1: A to B ---
        lrDX1  := stPointB[1] - stPointA[1];
        lrDY1  := stPointB[2] - stPointA[2];
        lrDTh1 := stPointB[3] - stPointA[3];
        lrL1   := MAX(0.001, SQRT(lrDX1*lrDX1 + lrDY1*lrDY1));
        
        // --- Line 2: B to C ---
        lrDX2  := stPointC[1] - stPointB[1];
        lrDY2  := stPointC[2] - stPointB[2];
        lrDTh2 := stPointC[3] - stPointB[3];
        lrL2   := MAX(0.001, SQRT(lrDX2*lrDX2 + lrDY2*lrDY2));
        
        // --- Line 3: C to A ---
        lrDX3  := stPointA[1] - stPointC[1];
        lrDY3  := stPointA[2] - stPointC[2];
        lrDTh3 := stPointA[3] - stPointC[3];
        lrL3   := MAX(0.001, SQRT(lrDX3*lrDX3 + lrDY3*lrDY3));

        // Reset Motion
        lrS_T   := 0;
        lrS_dot := 0;
        
        iCurrentSegment := 5; // Start with Approach
        GVL_MessageStaus.MessageStaus := 'Assistive: Guiding to Start Point A.';
        iState  := 5;


    // -----------------------------------------------------
    // STATE 5: APPROACH (Guiding Patient to Point A)
    // -----------------------------------------------------
    5:
        // A. Move the "Virtual Rabbit" along the path to A
        bAtPointA := UpdateTrapezoid(lrL_total := lrL_App);

        // B. Manually Calculate Setpoint (Interpolation)
        SetAppX     := lrApproachStartX + (lrDX_App / lrL_App) * lrS_T;
        SetAppY     := lrApproachStartY + (lrDY_App / lrL_App) * lrS_T;
        SetAppTheta := lrApproachStartTheta + (lrDTh_App / lrL_App) * lrS_T;
		
		SetVelAppX     := (lrDX_App / lrL_App) * lrS_dot;
        SetVelAppY     := (lrDY_App / lrL_App) * lrS_dot;
        SetVelAppTheta := (lrDTh_App / lrL_App) * lrS_dot;

        // C. Calculate Assistive Force (Spring/Damper)
        CalculateImpedanceForce(
            ActX := ActX, ActY := ActY, ActTheta := ActTheta,
            TargetX := SetAppX, TargetY := SetAppY, TargetTheta := SetAppTheta,
			 ActVelX := 0.0, ActVelY := 0.0, ActVelTheta := 0.0,  
			TargetVelX  := SetVelAppX, TargetVelY := SetVelAppY, TargetVelTheta := SetVelAppTheta, Fx_Cmd => CalcForces[1], 
            Fy_Cmd      => CalcForces[2], 
            MTheta_Cmd  => CalcForces[3] );

        // D. Convert to Torque & Drive
        JacobianTranspose(
            TargetFx := CalcForces[1], TargetFy := CalcForces[2], TargetMTheta := CalcForces[3],
            ActR := ActR, ActBeta := ActBeta,
            JointTorqueTarget => CalcTorques
        );

        DriveMotors(TorqueSetpoints := CalcTorques);

        // E. Check Completion
        IF bAtPointA THEN
            GVL_MessageStaus.MessageStaus  := 'Reached Point A. Resting...';
            bWaitEnable := TRUE; 
            iState := 7;
        END_IF


    // -----------------------------------------------------
    // STATE 7: WAIT (Rest at Corners)
    // -----------------------------------------------------
    7:
        // In Assistive mode, "Wait" means Zero Torque (Free Mode) 
        // or Holding Position (Stiff Mode). Here we use Zero Torque for rest.
        CalcTorques[1] := 0; 
        CalcTorques[2] := 0; 
        CalcTorques[3] := 0;
        DriveMotors(TorqueSetpoints := CalcTorques);

        IF fbWaitTimer.Q THEN
            bWaitEnable := FALSE;
            lrS_T   := 0;
            lrS_dot := 0;
            iCurrentSegment := 10; // Begin Main Triangle
            iState := 40;
            GVL_MessageStaus.MessageStaus  := 'Assistive: Path A to B started.';
        END_IF
		
(*


    // -----------------------------------------------------
    // STATE 10: MAIN ASSISTIVE LOOP (A->B->C->A)
    // -----------------------------------------------------
    10:
        // --- A. Select Target Segment Length ---
        CASE iCurrentSegment OF
            10: lrL_Target := lrL1; // A->B
            20: lrL_Target := lrL2; // B->C
            30: lrL_Target := lrL3; // C->A
        END_CASE

        // --- B. Move Virtual Target (The Rabbit) ---
        bSegmentDone := UpdateTrapezoid(lrL_total := lrL_Target);

        // --- C. Update Path Setpoints (Find X,Y of the Rabbit) ---
        // This method calculates SetX, SetY based on iCurrentSegment and lrS_T
        UpdatePathSetpoints(
            TargetX => SetX,
            TargetY => SetY,
            TargetTheta => SetTheta
        );

        // --- D. Calculate Impedance Force (The "Rubber Band") ---
        // Pulls the patient towards SetX/SetY
        CalculateImpedanceForce(
            ActX := ActX, ActY := ActY, ActTheta := ActTheta,
            TargetX := SetX, TargetY := SetY, TargetTheta := SetTheta,
            Kp_Cart := 0.5, // Stiffness: Adjust for "Assist Strength"
            Kd_Cart := 0.05, // Damping: Adjust for stability
            Fx_Cmd => CalcForces[1], 
            Fy_Cmd => CalcForces[2], 
            MTheta_Cmd => CalcForces[3]
        );

        // --- E. Convert Force to Torque ---
        JacobianTranspose(
            TargetFx := CalcForces[1], 
            TargetFy := CalcForces[2], 
            TargetMTheta := CalcForces[3],
            ActR := ActR, 
            ActBeta := ActBeta,
            JointTorqueTarget => CalcTorques
        );

        // --- F. Drive Motors ---
        DriveMotors(TorqueSetpoints := CalcTorques);

        // --- G. Segment Transition Logic ---
        IF bSegmentDone THEN
            bWaitEnable := TRUE; 
            lrS_T   := 0; // Reset Path Distance
            lrS_dot := 0; // Reset Velocity
        END_IF

        // Handle Waiting (Zero Torque during wait)
        IF bWaitEnable THEN
             // Optional: Zero torque to let patient rest arm
             CalcTorques[1] := 0; CalcTorques[2] := 0; CalcTorques[3] := 0;
             DriveMotors(TorqueSetpoints := CalcTorques);
        END_IF

        // Handle Timer Expiry & Switching
        IF fbWaitTimer.Q THEN
            bWaitEnable := FALSE;

            IF iCurrentSegment = 10 THEN
                iCurrentSegment := 20;
                GVL_MessageStaus.MessageStaus := 'Assistive: Path B to C.';
            ELSIF iCurrentSegment = 20 THEN
                iCurrentSegment := 30;
                GVL_MessageStaus.MessageStaus := 'Assistive: Path C to A.';
            ELSIF iCurrentSegment = 30 THEN
                iState := 40; // Done
                GVL_MessageStaus.MessageStaus := 'Assistive Task Complete.';
            END_IF
        END_IF
		
		*)

    // -----------------------------------------------------
    // STATE 40: FINISHED
    // -----------------------------------------------------
    40:
        bBusy := FALSE;
        // Zero Torque (Free Mode)
        CalcTorques[1] := 0; CalcTorques[2] := 0; CalcTorques[3] := 0;
        DriveMotors(TorqueSetpoints := CalcTorques);

END_CASE

METHOD CalculateImpedanceForce : BOOL
VAR_INPUT
    // --- Position Feedback (Where is the robot?) ---
    ActX     : LREAL; 
    ActY     : LREAL; 
    ActTheta : LREAL; 
    
    // --- Velocity Feedback (How fast is it moving?) ---
    // [CRITICAL] You must calculate this in your Main/Robot FB
    ActVelX     : LREAL;
    ActVelY     : LREAL;
    ActVelTheta : LREAL;

    // --- Targets (From Profile) ---
    TargetX     : LREAL;
    TargetY     : LREAL;
    TargetTheta : LREAL;
    
    // Optional: Target Velocity (Feedforward)
    // Set to 0.0 if you just want to hold a position
    TargetVelX     : LREAL := 0.0;
    TargetVelY     : LREAL := 0.0;
    TargetVelTheta : LREAL := 0.0;
    

    
END_VAR
VAR_OUTPUT
    // --- Final Force Commands ---
    Fx_Cmd      : LREAL;
    Fy_Cmd      : LREAL;
    MTheta_Cmd  : LREAL;
END_VAR
VAR
    // Errors
  //  Ex, Ey, ETheta    : LREAL; // Position Errors
    EvX, EvY, EvTheta : LREAL; // Velocity Errors
	
	Kp_Cart  : LREAL := 0.1 ; // Stiffness (N/mm) - "The Spring"
    Kd_Cart  : LREAL := 0.0; // Damping (Ns/mm)  - "The Honey"
    
    Kp_Rot   : LREAL := 0.05; // Rotational Stiffness
    Kd_Rot   : LREAL := 0.0; //tational Damping
END_VAR
// -----------------------------------------------------------------------------
// 1. Calculate Position Errors (The Spring Stretch)
// -----------------------------------------------------------------------------
Ex     := TargetX - ActX;
Ey     := TargetY - ActY;
ETheta := TargetTheta - ActTheta;

// -----------------------------------------------------------------------------
// 2. Calculate Velocity Errors (The Speed Difference)
// -----------------------------------------------------------------------------
// If TargetVel is 0, this becomes (0 - ActualVel), creating a braking force.
EvX     := TargetVelX - ActVelX;
EvY     := TargetVelY - ActVelY;
EvTheta := TargetVelTheta - ActVelTheta;

// -----------------------------------------------------------------------------
// 3. Apply Full Impedance Law: F = (Kp * PosError) + (Kd * VelError)
// -----------------------------------------------------------------------------
Fx_Cmd     := (Kp_Cart * Ex) + (Kd_Cart * EvX);
Fy_Cmd     := (Kp_Cart * Ey) + (Kd_Cart * EvY);
MTheta_Cmd := (Kp_Rot * ETheta) + (Kd_Rot * EvTheta);

CalculateImpedanceForce := TRUE;
END_METHOD

METHOD DriveMotors : BOOL
VAR_INPUT
	TorqueSetpoints : ARRAY [1..3] OF LREAL; // Calculated Torque (mNm)
END_VAR

VAR
	lrRatedTorque_Axis1 : LREAL := 810.425; 
    lrRatedTorque_Axis2 : LREAL := 383.934;
    lrRatedTorque_Axis3 : LREAL := 382.060;
	
END_VAR
// SCALING mm/s to Percentage
// Motor 1 (Axis 1)
lrTorqueSetpoint_Pct[1] := (TorqueSetpoints[1] / lrRatedTorque_Axis1) * 100.0;

// Motor 2 (Axis 2)
lrTorqueSetpoint_Pct[2] := (TorqueSetpoints[2] / lrRatedTorque_Axis2) * 100.0;

// Motor 3 (Axis 3)
lrTorqueSetpoint_Pct[3] := (TorqueSetpoints[3] / lrRatedTorque_Axis3) * 100.0;






fbTorqueAxis1(
    Axis             := GVL_Axes.Axis1,
    Execute          := TRUE,                 // Keep TRUE to stay active
    ContinuousUpdate := TRUE,                 // CRITICAL: Allows changing torque every cycle
    Torque           := lrTorqueSetpoint_Pct[1],   // Input from Jacobian
    Relative         := FALSE,  // Absolute Torque
	TorqueRamp         :=   1000.0,               
    VelocityLimitHigh:= MaxSpeedLimit,        // Safety: Prevent runaway if resistance is lost
    VelocityLimitLow := -MaxSpeedLimit
);

// -----------------------------------------------------------------------------
// AXIS 2 TORQUE CONTROL
// -----------------------------------------------------------------------------
fbTorqueAxis2(
    Axis             := GVL_Axes.Axis2,
    Execute          := TRUE,
    ContinuousUpdate := TRUE,
    Torque           := lrTorqueSetpoint_Pct[2],
    Relative         := FALSE,
	TorqueRamp         := 1000.0,
    VelocityLimitHigh:= MaxSpeedLimit,
    VelocityLimitLow := -MaxSpeedLimit
);

// -----------------------------------------------------------------------------
// AXIS 3 TORQUE CONTROL
// -----------------------------------------------------------------------------
fbTorqueAxis3(
    Axis             := GVL_Axes.Axis3,
    Execute          := TRUE,
    ContinuousUpdate := TRUE,
    Torque           := lrTorqueSetpoint_Pct[3],
    Relative         := FALSE,
	TorqueRamp         :=   1000.0,
    VelocityLimitHigh:= MaxSpeedLimit,
    VelocityLimitLow := -MaxSpeedLimit
);

DriveMotors := TRUE;
END_METHOD

METHOD JacobianTranspose : BOOL
VAR_INPUT
    // Inputs (Forces & Robot State)
    TargetFx     : LREAL; // Force in X (N)
    TargetFy     : LREAL; // Force in Y (N)
    TargetMTheta : LREAL; // Moment for Wrist (Nmm)
    
    ActR         : LREAL; // Current Radius (mm)
    ActBeta      : LREAL; // Current Arm Angle (Degrees) - Corresponds to 'Beta'
END_VAR
VAR_OUTPUT
    // Outputs (Motor Torques)
    JointTorqueTarget : ARRAY [1..3] OF LREAL;
END_VAR
VAR
    // Local Variables
    BetaRad : LREAL;
    R_mm    : LREAL;
    PI_180    : LREAL := 0.0174532925199433; 
    // Jacobian Matrix Elements
    J11, J12, J13 : LREAL;
    J21, J22, J23 : LREAL;
    J31, J32, J33 : LREAL;
END_VAR
// -----------------------------------------------------------------------------
// 1. Assign local values (Consistent with your Inverse Jacobian style)
// -----------------------------------------------------------------------------
BetaRad := ActBeta * PI_180; // Convert Degree to Radian
R_mm    := ActR;

// -----------------------------------------------------------------------------
// 2. Populate Jacobian Matrix Elements (Derived from your Forward Kinematics)
// -----------------------------------------------------------------------------
// Row 1: How X changes with motors
J11 := -R_mm * GVL_ConstantCoefficent.K1 * PI_180 * COS(BetaRad); 
J12 :=  GVL_ConstantCoefficent.K2 * SIN(BetaRad);
J13 := -GVL_ConstantCoefficent.K2 * SIN(BetaRad);

// Row 2: How Y changes with motors
J21 :=  R_mm * GVL_ConstantCoefficent.K1 * PI_180 * SIN(BetaRad);
J22 :=  GVL_ConstantCoefficent.K2 * COS(BetaRad);
J23 := -GVL_ConstantCoefficent.K2 * COS(BetaRad);

// Row 3: How Theta (Wrist) changes with motors
J31 := 0.0;
J32 := -GVL_ConstantCoefficent.K3 / 2.0;
J33 := -GVL_ConstantCoefficent.K3 / 2.0;

// -----------------------------------------------------------------------------
// 3. Apply Jacobian Transpose (Tau = J_Transpose * Force)
// -----------------------------------------------------------------------------

// Motor 1 Torque: Sum of (Col 1 * Forces)
JointTorqueTarget[1] := (J11 * TargetFx) + (J21 * TargetFy) + (J31 * TargetMTheta);

// Motor 2 Torque: Sum of (Col 2 * Forces)
JointTorqueTarget[2] := (J12 * TargetFx) + (J22 * TargetFy) + (J32 * TargetMTheta);

// Motor 3 Torque: Sum of (Col 3 * Forces)
JointTorqueTarget[3] := (J13 * TargetFx) + (J23 * TargetFy) + (J33 * TargetMTheta);

JacobianTranspose := TRUE;
END_METHOD

METHOD UpdatePathSetpoints : BOOL
VAR_INPUT
END_VAR

CASE iCurrentSegment OF
    10: // Line A -> B
        IF lrL1 > 0.0 THEN
            stCurrentSet[1] := stPointA[1] + (lrDX1 / lrL1) * lrS_T;
            stCurrentSet[2] := stPointA[2] + (lrDY1 / lrL1) * lrS_T;
            stCurrentSet[3] := stPointA[3] + (lrDTh1 / lrL1) * lrS_T;
            
            // Calculate Feedforward Velocities (Unit Vector * Current Speed)
            lrVx_FF := (lrDX1 / lrL1) * lrS_dot;
            lrVy_FF := (lrDY1 / lrL1) * lrS_dot;
            lrVTh_FF := (lrDTh1 / lrL1) * lrS_dot;
        END_IF;

    20: // Line B -> C
        IF lrL2 > 0.0 THEN
            stCurrentSet[1] := stPointB[1] + (lrDX2 / lrL2) * lrS_T;
            stCurrentSet[2] := stPointB[2] + (lrDY2 / lrL2) * lrS_T;
            stCurrentSet[3] := stPointB[3] + (lrDTh2 / lrL2) * lrS_T;
            
            lrVx_FF := (lrDX2 / lrL2) * lrS_dot;
            lrVy_FF := (lrDY2 / lrL2) * lrS_dot;
            lrVTh_FF := (lrDTh2 / lrL2) * lrS_dot;
        END_IF;

    30: // Line C -> A
        IF lrL3 > 0.0 THEN
            stCurrentSet[1] := stPointC[1] + (lrDX3 / lrL3) * lrS_T;
            stCurrentSet[2] := stPointC[2] + (lrDY3 / lrL3) * lrS_T;
            stCurrentSet[3] := stPointC[3] + (lrDTh3 / lrL3) * lrS_T;
            
            lrVx_FF := (lrDX3 / lrL3) * lrS_dot;
            lrVy_FF := (lrDY3 / lrL3) * lrS_dot;
            lrVTh_FF := (lrDTh3 / lrL3) * lrS_dot;
        END_IF;
END_CASE
END_METHOD

METHOD UpdateTrapezoid : BOOL
VAR_INPUT
	lrL_total : LREAL;
	
END_VAR

VAR
		
    dist_rem  : LREAL;
    CycleTime : LREAL := 0.01;  //plc cycle time is 10 ms
	S_dec : LREAL; // calcullated stopping distance
	
END_VAR
// This method calculates the current velocity and distance scalar for the move.

s_dec := (lrVmax * lrVmax) / (2.0 * lrAcc);
dist_rem := lrL_total - lrS_T;

IF dist_rem > s_dec THEN
    lrS_dot := MIN(lrS_dot + (lrAcc * CycleTime), lrVmax);
ELSE
    lrS_dot := SQRT(2.0 * lrAcc * MAX(0.0, dist_rem));
END_IF

lrS_T := lrS_T + (lrS_dot * CycleTime);

IF dist_rem <= 0.001 THEN
    UpdateTrapezoid := TRUE; // Signal segment complete
END_IF
END_METHOD

END_FUNCTION_BLOCK

// ---- POUs/FB_AdmittanceController.TcPOU
FUNCTION_BLOCK FB_AdmittanceController
VAR_INPUT
	
END_VAR
VAR_OUTPUT
END_VAR
VAR
END_VAR

END_FUNCTION_BLOCK

// ---- POUs/FB_ForceController.TcPOU
FUNCTION_BLOCK FB_ForceController
VAR_INPUT
END_VAR
VAR_OUTPUT
END_VAR
VAR
END_VAR

END_FUNCTION_BLOCK

// ---- POUs/FB_DynamicsCompensator.TcPOU
FUNCTION_BLOCK FB_DynamicsCompensator
VAR_INPUT
	// 1. Feature Flags (Explicit and isolated)
    EnableFrictionComp : BOOL;       
    EnableInertiaComp  : BOOL;
	
	// Kinematic data
	
END_VAR
VAR_OUTPUT
	TotalCompTorque    : ST_JointTorque;
END_VAR
VAR
	CalculatedFriction : ST_JointTorque;
    CalculatedInertia  : ST_JointTorque;
END_VAR

// 1. FRICTION COMPENSATION
IF EnableFrictionComp THEN
    //
ELSE
    CalculatedFriction.M1 := 0.0;
    CalculatedFriction.M2 := 0.0;
    CalculatedFriction.M3 := 0.0;
END_IF

// 2. INERTIA COMPENSATION
IF EnableInertiaComp THEN
    //
ELSE
    CalculatedInertia.M1 := 0.0;
    CalculatedInertia.M2 := 0.0;
    CalculatedInertia.M3 := 0.0;
END_IF

// 3. COMBINE FOR OUTPUT
TotalCompTorque.M1 := CalculatedFriction.M1 + CalculatedInertia.M1;
TotalCompTorque.M2 := CalculatedFriction.M2 + CalculatedInertia.M2;
TotalCompTorque.M3 := CalculatedFriction.M3 + CalculatedInertia.M3;

END_FUNCTION_BLOCK

// ---- POUs/FB_VirtuallWall.TcPOU
FUNCTION_BLOCK FB_VirtuallWall
VAR_INPUT
	bEnable     : BOOL ;     // Enable Virtual Wall Controller
    Endeffectorstatus : ST_CartesianState;
    fStiffness  : LREAL := 0.06;     // Virtual Wall Stiffness K [N/mm]
    fDamping    : LREAL := 0.01;    // Virtual Wall Damping B [N/(mm/s)]
	WallSetPointXandY : ARRAY[1..4, 1..2] OF LREAL ;
END_VAR
VAR_OUTPUT
	WallCartesianForce : ST_CartesianForces;
	bInContact  : BOOL;
END_VAR
VAR
	// Pre-calculated geometric constant for slanted lines: SQRT(157^2 + 150^2)
    cNorm23     : LREAL := 217.138209447043; 

    // walls Position
	TopWall_Constant : LREAL  := 260.0; //  y =Constant   This number is predefined walls if set new upperside wall it will change
	BottomWall_Constant : LREAL  := -10.0; // Bottom Wall (y = Constant) This number is predefined walls if set new upperside wall it will change
	RightWall_A : LREAL; // Ax+By + C=0 for right wall
	RightWall_B : LREAL;  // Ax+By + C =0for right wall
	RightWall_C : LREAL;  // Ax+By + C=0 for right wall
	
	LeftWall_A : LREAL; // Ax+By + C =0 for Left wall 
	LeftWall_B : LREAL; // Ax+By + C=0 for Left wall
	LeftWall_C : LREAL; // Ax+By + C =0 for Left wall
	
	
    NormTop      : ARRAY[1..2] OF LREAL := [ 0.0, -1.0];             // Top Wall (y = 260)
    
    NormBottom      : ARRAY[1..2] OF LREAL := [ 0.0,  1.0];             // Bottom Wall (y = -10)

  // Calculation Virtuall Wall 
  x_COR_CartezianforCalculationRightLeftWall : LREAL := 0.0; //Center of rotation in cartezian (x=0 y=)
  y_COR_CartezianforCalculationRightLeftWall : LREAL := 464.0;  //Center of rotation in cartezian (x=0 y=)
  y_SetwallRightWall : LREAL;
  x_SetwallRightWall : LREAL;
  y_SetwallLeftWall : LREAL;
  x_SetwallLeftWall : LREAL;
  RightWall_NormalMagnitude : LREAL;
  NormRight     : ARRAY[1..2] OF LREAL;  // Right Wall
  LeftWall_NormalMagnitude : LREAL;
  NormLeft     : ARRAY[1..2] OF LREAL;  // Left Wall


// Calculation Variables
    fDelta      : LREAL;            // Penetration depth [mm]
    fVnormal    : LREAL;            // Velocity along inward normal [mm/s]
    fDampEff    : LREAL;            // Non-sticky effective damping force
    fForceMag   : LREAL;            // Force magnitude for individual wall
	
	///
	fForceX     : LREAL;            // Virtual Wall Restoring Force X [N]
    fForceY     : LREAL;            // Virtual Wall Restoring Force Y [N]
                 // TRUE if penetrating any boundary
	fActY: LREAL;
	fActX: LREAL;
	fActXdot: LREAL;
	fActYdot: LREAL;
	fbRobotKinematicForJacobianInverse : FB_RobotKinematics;
	WallJointState : ST_JointState;
	
//	JointData_Transed: INT;
 
END_VAR

TopWall_Constant := WallSetPointXandY[1,2];
BottomWall_Constant := WallSetPointXandY [2,2];
x_SetwallRightWall := WallSetPointXandY [3,1];
y_SetwallRightWall :=  WallSetPointXandY [3,2];
x_SetwallLeftWall := WallSetPointXandY [4,1];
y_SetwallLeftWall := WallSetPointXandY [4,2];

// Reset outputs at start of cycle
fForceX := 0.0;
fForceY := 0.0;
bInContact := FALSE;


// Right wall equation: A*x + B*y + C = 0

RightWall_A :=
    y_COR_CartezianforCalculationRightLeftWall - y_SetwallRightWall;

RightWall_B :=
    x_SetwallRightWall - x_COR_CartezianforCalculationRightLeftWall;

RightWall_C :=
    (x_COR_CartezianforCalculationRightLeftWall * y_SetwallRightWall)
    - (x_SetwallRightWall * y_COR_CartezianforCalculationRightLeftWall);


// UnitNormal of Right wall

RightWall_NormalMagnitude := SQRT(
    RightWall_A * RightWall_A +
    RightWall_B * RightWall_B
);

IF RightWall_NormalMagnitude > 0.001 THEN
    NormRight[1] := -RightWall_A / RightWall_NormalMagnitude;
    NormRight[2] := -RightWall_B / RightWall_NormalMagnitude;
ELSE
    NormRight[1] := 0.0;
    NormRight[2] := 0.0;
END_IF;



// Left wall equation: A*x + B*y + C = 0

LeftWall_A :=
    y_COR_CartezianforCalculationRightLeftWall - y_SetwallLeftWall;

LeftWall_B :=
    x_SetwallLeftWall - x_COR_CartezianforCalculationRightLeftWall;

LeftWall_C :=
    (x_COR_CartezianforCalculationRightLeftWall * y_SetwallLeftWall)
    - (x_SetwallLeftWall * y_COR_CartezianforCalculationRightLeftWall);
	
	// UnitNormal of Left wall

LeftWall_NormalMagnitude := SQRT(
    LeftWall_A * LeftWall_A +
    LeftWall_B * LeftWall_B
);

IF LeftWall_NormalMagnitude > 0.001 THEN
    NormLeft[1] := LeftWall_A / LeftWall_NormalMagnitude;
    NormLeft[2] := LeftWall_B / LeftWall_NormalMagnitude;
ELSE
    NormLeft[1] := 0.0;
    NormLeft[2] := 0.0;
END_IF;


// 

fActX := Endeffectorstatus.Position.X;
fActY := Endeffectorstatus.Position.Y;
fActXdot := Endeffectorstatus.Velocity.Vx;
fActYdot := Endeffectorstatus.Velocity.Vy;


WallCartesianForce.Fx := 0.0;
WallCartesianForce.Fy := 0.0;
WallCartesianForce.Mtheta := 0.0;


IF NOT bEnable THEN
    RETURN;
END_IF;





// -------------------------------------------------------------
// LINE 1: Top Wall 
// -------------------------------------------------------------
fDelta := fActY - TopWall_Constant; 
IF fDelta > 0.0 THEN
    bInContact := TRUE;
    fVnormal := (fActXdot * NormTop[1]) + (fActYdot * NormTop[2]);
    
    // Apply damping only when moving deeper into the wall
    IF fVnormal < 0.0 THEN
        fDampEff := -fDamping * fVnormal;
    ELSE
        fDampEff := 0.0;
    END_IF;
    
    fForceMag := (fStiffness * fDelta) + fDampEff;
    fForceX := fForceX + (fForceMag * NormTop[1]);
    fForceY := fForceY + (fForceMag * NormTop[2]);
END_IF;

// -------------------------------------------------------------
// LINE 2: RIGHT WALL (Ax + By + C = 0)
// -------------------------------------------------------------

IF RightWall_NormalMagnitude > 0.001 THEN

    fDelta := (
        RightWall_A * fActX +
        RightWall_B * fActY +
        RightWall_C
    ) / RightWall_NormalMagnitude;

    IF fDelta > 0.0 THEN

        bInContact := TRUE;

        fVnormal :=
            (fActXdot * NormRight[1]) +
            (fActYdot * NormRight[2]);

        // Apply damping only when moving deeper into the wall
        IF fVnormal < 0.0 THEN
            fDampEff := -fDamping * fVnormal;
        ELSE
            fDampEff := 0.0;
        END_IF;

        fForceMag := (fStiffness * fDelta) + fDampEff;

        fForceX := fForceX + (fForceMag * NormRight[1]);
        fForceY := fForceY + (fForceMag * NormRight[2]);

    END_IF;

END_IF;


// -------------------------------------------------------------
// LINE 3: LEFT WALL (Ax + By + C = 0)
// -------------------------------------------------------------

IF LeftWall_NormalMagnitude > 0.001 THEN

    fDelta := -(
        LeftWall_A * fActX +
        LeftWall_B * fActY +
        LeftWall_C
    ) / LeftWall_NormalMagnitude;

    IF fDelta > 0.0 THEN

        bInContact := TRUE;

        fVnormal :=
            (fActXdot * NormLeft[1]) +
            (fActYdot * NormLeft[2]);

        // Apply damping only when moving deeper into the wall
        IF fVnormal < 0.0 THEN
            fDampEff := -fDamping * fVnormal;
        ELSE
            fDampEff := 0.0;
        END_IF;

        fForceMag := (fStiffness * fDelta) + fDampEff;

        fForceX := fForceX + (fForceMag * NormLeft[1]);
        fForceY := fForceY + (fForceMag * NormLeft[2]);

    END_IF;

END_IF;

// -------------------------------------------------------------
// LINE 4: Bottom Wall (y = -10 mm)
// -------------------------------------------------------------


fDelta := BottomWall_Constant - fActY;

IF fDelta > 0.0 THEN

    bInContact := TRUE;

    fVnormal :=
        (fActXdot * NormBottom[1]) +
        (fActYdot * NormBottom[2]);

    IF fVnormal < 0.0 THEN
        fDampEff := -fDamping * fVnormal;
    ELSE
        fDampEff := 0.0;
    END_IF;

    fForceMag := (fStiffness * fDelta) + fDampEff;

    fForceX := fForceX + (fForceMag * NormBottom[1]);
    fForceY := fForceY + (fForceMag * NormBottom[2]);

END_IF;

 GVL_HMI.VirtualWallContact := bInContact;
WallCartesianForce.Fx := fForceX;
 WallCartesianForce.Fy := fForceY;
 WallCartesianForce.Mtheta := 0.0; // wrist

END_FUNCTION_BLOCK

// ---- POUs/FB_DriveInterface.TcPOU
FUNCTION_BLOCK FB_DriveInterface
VAR_INPUT
TorqueSetpoints : ST_JointTorque;
Config           : ST_TherapyConfig;
END_VAR
VAR_OUTPUT
END_VAR
VAR
	
	lrRatedTorque_Axis1 : LREAL := 810.425; 
    lrRatedTorque_Axis2 : LREAL := 383.934;
    lrRatedTorque_Axis3 : LREAL := 382.060;
	
	fbTorqueAxis1    : MC_TorqueControl;
    fbTorqueAxis2    : MC_TorqueControl;
    fbTorqueAxis3    : MC_TorqueControl;
	lrTorqueSetpoint_Pct : ST_JointTorque;
	
	lrEffectiveSpeedHigh  : LREAL;
    lrEffectiveSpeedLow   : LREAL;
	ErrorAxisA: BOOL;
	ErrorAxisID: UDINT;
	Execute_A : BOOL ;
	Execute_B : BOOL ;
	Execute_C : BOOL ;
	TurnOnMotors: BOOL := FALSE;
	
	
	ErrorAxisID_A: UDINT;
	ErrorAxisID_B: UDINT;
	ErrorAxisB: BOOL;
	ErrorAxisC: BOOL;
	ErrorAxisID_C: UDINT;
	torqueofaxisB: BOOL;
	BisBusy: BOOL;
	BisActive: BOOL;
	torqueofaxisA: BOOL;
	AisBusy: BOOL;
	AisActive: BOOL;
END_VAR

// 1. Clamp Positive Game Limit between 0.0 and +GlobalVelocityLimit
lrEffectiveSpeedHigh := LIMIT(
    0.0, 
    ABS(Config.GlobalVelocityLimit), // THIS Data should changed based on game currently I put equal tp g;pbalspeedlimitHigh
    ABS(Config.GlobalVelocityLimit)
);

// 2. Clamp Negative Game Limit between -GlobalVelocityLimit and 0.0
lrEffectiveSpeedLow  := LIMIT(
    -ABS(Config.GlobalVelocityLimit), // THIS Data should changed based on game currently I put equal tp g;pbalspeedlimitHigh
    -ABS(Config.GlobalVelocityLimit), 
    0.0
);



// SCALING NM to Percentage
// Motor 1 (Axis 1)
lrTorqueSetpoint_Pct.M1 := (TorqueSetpoints.M1 / lrRatedTorque_Axis1) * 100.0;

// Motor 2 (Axis 2)
lrTorqueSetpoint_Pct.M2 := (TorqueSetpoints.M2 / lrRatedTorque_Axis2) * 100.0;
// Motor 3 (Axis 3)
lrTorqueSetpoint_Pct.M3 := (TorqueSetpoints.M3 / lrRatedTorque_Axis3) * 100.0;

lrTorqueSetpoint_Pct.M1 := TorqueSetpoints.M1;
lrTorqueSetpoint_Pct.M2 := TorqueSetpoints.M2;
lrTorqueSetpoint_Pct.M3 := TorqueSetpoints.M3;


// lrTorqueSetpoint_Pct.M1 := 20.0;
// lrTorqueSetpoint_Pct.M2 := 50.0;
// lrTorqueSetpoint_Pct.M3 := -50.0;	

//lrTorqueSetpoint_Pct.M1 := TorqueSetpoints.M1;
//lrTorqueSetpoint_Pct.M2 := TorqueSetpoints.M2;
//lrTorqueSetpoint_Pct.M3 := TorqueSetpoints.M3;

Execute_A := GVL_HMI.ContinueTOWorkspaceLimits;
Execute_B := GVL_HMI.ContinueTOWorkspaceLimits;
Execute_C := GVL_HMI.ContinueTOWorkspaceLimits;


fbTorqueAxis1(
    Axis             := GVL_Axes.Axis1,
    Execute          := Execute_A,                 // Keep TRUE to stay active
    ContinuousUpdate := TRUE,                 // CRITICAL: Allows changing torque every cycle
    Torque           := lrTorqueSetpoint_Pct.M1,   // Input from Jacobian
    Relative         := FALSE,  // Absolute Torque
	TorqueRamp         :=   100.0,               
    VelocityLimitHigh:= lrEffectiveSpeedHigh,        // Safety: Prevent runaway if resistance is lost
    VelocityLimitLow := lrEffectiveSpeedLow,
	InTorque => torqueofaxisA,
	Busy=> AisBusy,
	Active => AisActive,
	Error => ErrorAxisA ,
	ErrorID => ErrorAxisID_A
);

// -----------------------------------------------------------------------------
// AXIS 2 TORQUE CONTROL
// -----------------------------------------------------------------------------
fbTorqueAxis2(
    Axis             := GVL_Axes.Axis2,
    Execute          := Execute_B,
    ContinuousUpdate := TRUE,
    Torque           := lrTorqueSetpoint_Pct.M2,
    Relative         := FALSE,
	TorqueRamp         := 100.0,
    VelocityLimitHigh:= lrEffectiveSpeedHigh,        // Safety: Prevent runaway if resistance is lost
    VelocityLimitLow := lrEffectiveSpeedLow,
	InTorque => torqueofaxisB,
	Busy=> BisBusy,
	Active => BisActive,
	
	Error => ErrorAxisB ,
	ErrorID => ErrorAxisID_B
);

// -----------------------------------------------------------------------------
// AXIS 3 TORQUE CONTROL
// -----------------------------------------------------------------------------
fbTorqueAxis3(
    Axis             := GVL_Axes.Axis3,
    Execute          := Execute_C,
    ContinuousUpdate := TRUE,
    Torque           := lrTorqueSetpoint_Pct.M3,
    Relative         := FALSE,
	TorqueRamp         :=   100.0,
    VelocityLimitHigh:= lrEffectiveSpeedHigh,        // Safety: Prevent runaway if resistance is lost
    VelocityLimitLow := lrEffectiveSpeedLow,
	Error => ErrorAxisC,
	ErrorID => ErrorAxisID_C
);

// DriveMotors := TRUE;

END_FUNCTION_BLOCK

// ---- POUs/HMI_FunBlock/FB_HMI_TherapyConfiguration.TcPOU
FUNCTION_BLOCK FB_HMI_TherapyConfiguration
VAR_INPUT
	CartesianDataTransedFromJointSpace : ST_CartesianState;
END_VAR
VAR_OUTPUT
	 WallSetPointXandY : ARRAY[1..4, 1..2] OF LREAL := [
    0.0, 370.408,        // Top wall
    0.0, -12.245,        // Bottom wall
    168.367, 370.408,    // Right wall
    -168.367, 370.408    // Left wall
];
END_VAR
VAR
sPolygonPoints: STRING(255);
ActiveWall: INT;
EndEffectorPixcelPosY : INT;
EndEffectorPixcelPosX : INT;

//
// ActiveWall: INT:=1;
	X_A : INT ;
	Y_AB : INT ;
	X_B : INT ;
	
	X_C : INT ;
	Y_CD : INT ;
	X_D: INT ;
	nLength: INT;
	
	X_ConstantoFRotationalCenterPixcel : INT := 260;
Y_ConstantoFRotationalCenterPixcel : INT := -60;

bPolygonInitialized: BOOL;
(* Set button edge *)
bSetWall : BOOL;
bSetWallOld : BOOL;
bSetWallRisingEdge : BOOL;

//
fbSetWallTrig : R_TRIG;

    fbTopWallTrig : R_TRIG;
    fbBottomWallTrig : R_TRIG;
    fbRightWallTrig : R_TRIG;
    fbLeftWallTrig : R_TRIG;

// WRIST VARIABLE
// =========================================================
// WRIST PURPLE LINE
// =========================================================

fWristLineX : LREAL;                 // X of moving endpoint
fWristLineY : LREAL;                 // Y of moving endpoint

fWristCenterX : LREAL := 100.0;      // Fixed center X [pixel]
fWristCenterY : LREAL := 100.0;      // Fixed center Y [pixel]
fWristRadius  : LREAL := 100.0;      // Purple line length [pixel]

fAngleRad : LREAL;                   // Wrist angle [rad]


// =========================================================
// WRIST VIRTUAL WALL
// =========================================================

// 0 = No wall active
// 1 = Right wall active
// 2 = Left wall active
WristWall : INT := 0;

// Polygon:
// [1,*] = A
// [2,*] = B
// [3,*] = C
aWristPolygon : ARRAY[1..3, 1..2] OF LREAL;

// Polygon string for HMI binding
sWristPolygonPoints : STRING(255);


// =========================================================
// SET / SAVE
// =========================================================

bWristPolygonInitialized : BOOL := FALSE;

bWristSetOld : BOOL := FALSE;
bWristSetRisingEdge : BOOL;

bWristSetEnable : BOOL;
bWristWallInvalid : BOOL;

// 
fbRightWristWallTrig : R_TRIG;
    fbLeftWristWallTrig  : R_TRIG;
    fbWristSetTrig       : R_TRIG;

   // bWristSetRisingEdge  : BOOL;
END_VAR

GVL_HMI.CurrentTherapyConfig.ControllerType := E_ControllerType.ControlNone;
GVL_HMI.CurrentTherapyConfig.GlobalVelocityLimit := 100;

IF GVL_HMI.EableVirtuallWall_Planar THEN
	
PlanarHMIWall();

END_IF



WristHMIWall();
ButtonStatus();

nLength := LEN(sPolygonPoints);

METHOD ButtonStatus 
VAR
  
END_VAR
IF NOT GVL_HMI.bActiveMode
   AND NOT GVL_HMI.bPassiveMode
   AND NOT GVL_HMI.bAssistiveMode
   AND NOT GVL_HMI.bResistiveMode
   AND NOT GVL_HMI.bGameBasedMode THEN

    // Default mode
    GVL_HMI.bGameBasedMode := TRUE;

END_IF;
END_METHOD

METHOD PlanarHMIWall : BOOL
VAR_INPUT
END_VAR

VAR
	
	


LineRight_Y : LREAL;
LineRight_X : LREAL;
EndEffectorLocalX : INT;
EndEffectorLocalY : INT;
	
	LineLeft_Y: LREAL;
	LineLeft_X: LREAL;
	
	aPolygon : ARRAY[1..4, 1..2] OF INT;
	i: INT;
	
	DeltaY: INT;
END_VAR
(************************************************************
    WALL SELECTION
    Select a new wall ONLY when no wall is currently active
*************************************************************)

fbTopWallTrig(
    CLK := GVL_HMI.TopPlanarWall_But
);

fbBottomWallTrig(
    CLK := GVL_HMI.BottomPlanarWall_But
);

fbRightWallTrig(
    CLK := GVL_HMI.RightPlanarWall_But
);

fbLeftWallTrig(
    CLK := GVL_HMI.LeftPlanarWall_But
);


IF ActiveWall = 0 THEN

    IF fbTopWallTrig.Q THEN

        ActiveWall := 1;

    ELSIF fbBottomWallTrig.Q THEN

        ActiveWall := 2;

    ELSIF fbRightWallTrig.Q THEN

        ActiveWall := 3;

    ELSIF fbLeftWallTrig.Q THEN

        ActiveWall := 4;

    END_IF;

END_IF;


(************************************************************
    INITIALIZE POLYGON ONLY ONCE
*************************************************************)

IF NOT bPolygonInitialized THEN

    X_A := 150;
    Y_AB := 10;
    X_B := 370;

    X_C := 765;
    Y_CD := 260;
    X_D := -245;

    bPolygonInitialized := TRUE;

END_IF;


(************************************************************
    GET END-EFFECTOR POSITION
*************************************************************)

EndEffectorPixcelPosX :=
    GVL_HMI.EndeffectorPositionPixcelUnit_X;

EndEffectorPixcelPosY :=
    GVL_HMI.EndeffectorPositionPixcelUnit_Y;


(************************************************************
    CONVERT TO POLYGON COORDINATE SYSTEM
*************************************************************)

EndEffectorLocalX :=
    EndEffectorPixcelPosX - 233;

EndEffectorLocalY :=
    EndEffectorPixcelPosY - 443 + 15;


(************************************************************
    SET BUTTON RISING EDGE
*************************************************************)

fbSetWallTrig(
    CLK := GVL_HMI.SETPlanarWall_But
);

bSetWallRisingEdge := fbSetWallTrig.Q;


(************************************************************
    MODIFY ACTIVE WALL ONLY WHILE SET IS NOT PRESSED
*************************************************************)

IF ActiveWall <> 0 THEN

    CASE ActiveWall OF


        (********************************************************
            1: TOP WALL AB
        *********************************************************)

        1:

             Y_AB := EndEffectorLocalY;


    (* Point A:
       line AD passes through rotation center R *)
    X_A := LREAL_TO_INT(

        TO_LREAL(X_ConstantoFRotationalCenterPixcel)

        +

        (
            TO_LREAL(150)
            -
            TO_LREAL(X_ConstantoFRotationalCenterPixcel)
        )

        *

        (
            TO_LREAL(Y_AB)
            -
            TO_LREAL(Y_ConstantoFRotationalCenterPixcel)
        )

        /

        (
            TO_LREAL(10)
            -
            TO_LREAL(Y_ConstantoFRotationalCenterPixcel)
        )

    );


    (* Point B:
       line BC passes through rotation center R *)
    X_B := LREAL_TO_INT(

        TO_LREAL(X_ConstantoFRotationalCenterPixcel)

        +

        (
            TO_LREAL(370)
            -
            TO_LREAL(X_ConstantoFRotationalCenterPixcel)
        )

        *

        (
            TO_LREAL(Y_AB)
            -
            TO_LREAL(Y_ConstantoFRotationalCenterPixcel)
        )

        /

        (
            TO_LREAL(10)
            -
            TO_LREAL(Y_ConstantoFRotationalCenterPixcel)
        )

    );


        (********************************************************
            2: BOTTOM WALL DC
        *********************************************************)

        2:

            DeltaY :=
                EndEffectorLocalY - Y_CD;

            X_D := REAL_TO_INT(
                INT_TO_REAL(X_D)
                +
                INT_TO_REAL(DeltaY)
                * (-395.0 / 250.0)
            );

            X_C := REAL_TO_INT(
                INT_TO_REAL(X_C)
                +
                INT_TO_REAL(DeltaY)
                * (395.0 / 250.0)
            );

            Y_CD :=
                EndEffectorLocalY;


        (********************************************************
            3: RIGHT WALL BC
        *********************************************************)

        3:

            X_B := LREAL_TO_INT(

                TO_LREAL(X_ConstantoFRotationalCenterPixcel)

                +

                (
                    TO_LREAL(EndEffectorLocalX)
                    -
                    TO_LREAL(X_ConstantoFRotationalCenterPixcel)
                )

                *

                (
                    TO_LREAL(Y_AB)
                    -
                    TO_LREAL(Y_ConstantoFRotationalCenterPixcel)
                )

                /

                (
                    TO_LREAL(EndEffectorLocalY)
                    -
                    TO_LREAL(Y_ConstantoFRotationalCenterPixcel)
                )

            );


            X_C := LREAL_TO_INT(

                TO_LREAL(X_ConstantoFRotationalCenterPixcel)

                +

                (
                    TO_LREAL(EndEffectorLocalX)
                    -
                    TO_LREAL(X_ConstantoFRotationalCenterPixcel)
                )

                *

                (
                    TO_LREAL(Y_CD)
                    -
                    TO_LREAL(Y_ConstantoFRotationalCenterPixcel)
                )

                /

                (
                    TO_LREAL(EndEffectorLocalY)
                    -
                    TO_LREAL(Y_ConstantoFRotationalCenterPixcel)
                )

            );


        (********************************************************
            4: LEFT WALL AD
        *********************************************************)

        4:

            X_A := LREAL_TO_INT(

                TO_LREAL(X_ConstantoFRotationalCenterPixcel)

                +

                (
                    TO_LREAL(EndEffectorLocalX)
                    -
                    TO_LREAL(X_ConstantoFRotationalCenterPixcel)
                )

                *

                (
                    TO_LREAL(Y_AB)
                    -
                    TO_LREAL(Y_ConstantoFRotationalCenterPixcel)
                )

                /

                (
                    TO_LREAL(EndEffectorLocalY)
                    -
                    TO_LREAL(Y_ConstantoFRotationalCenterPixcel)
                )

            );


            X_D := LREAL_TO_INT(

                TO_LREAL(X_ConstantoFRotationalCenterPixcel)

                +

                (
                    TO_LREAL(EndEffectorLocalX)
                    -
                    TO_LREAL(X_ConstantoFRotationalCenterPixcel)
                )

                *

                (
                    TO_LREAL(Y_CD)
                    -
                    TO_LREAL(Y_ConstantoFRotationalCenterPixcel)
                )

                /

                (
                    TO_LREAL(EndEffectorLocalY)
                    -
                    TO_LREAL(Y_ConstantoFRotationalCenterPixcel)
                )

            );

    END_CASE;

END_IF;


(************************************************************
    WHEN SET IS PRESSED, FIX THE WALL
*************************************************************)
IF bSetWallRisingEdge THEN

    CASE ActiveWall OF

        // TOP WALL AB
        1:
            WallSetPointXandY[1,1] := 0.0;
			WallSetPointXandY[1,2] := CartesianDataTransedFromJointSpace.Position.Y;
                


        // BOTTOM WALL DC
        2:
            WallSetPointXandY[2,1] := 0.0;
			WallSetPointXandY[2,2] := CartesianDataTransedFromJointSpace.Position.Y;


        // RIGHT WALL BC
        3:
            WallSetPointXandY[3,1] :=CartesianDataTransedFromJointSpace.Position.X;
			WallSetPointXandY[3,2] := CartesianDataTransedFromJointSpace.Position.Y;


        // LEFT WALL AD
        4:
            WallSetPointXandY[4,1] :=CartesianDataTransedFromJointSpace.Position.X;
			WallSetPointXandY[4,2] := CartesianDataTransedFromJointSpace.Position.Y;

    END_CASE;


    // No wall is currently being edited
    ActiveWall := 0;

    // Reset SET button
    GVL_HMI.SETPlanarWall_But := FALSE;

    // Deselect all wall buttons
    GVL_HMI.TopPlanarWall_But := FALSE;
    GVL_HMI.BottomPlanarWall_But := FALSE;
    GVL_HMI.RightPlanarWall_But := FALSE;
    GVL_HMI.LeftPlanarWall_But := FALSE;

END_IF;


(************************************************************
    UPDATE POLYGON ARRAY
*************************************************************)

aPolygon[1, 1] := X_A;
aPolygon[1, 2] := Y_AB;

aPolygon[2, 1] := X_B;
aPolygon[2, 2] := Y_AB;

aPolygon[3, 1] := X_C;
aPolygon[3, 2] := Y_CD;

aPolygon[4, 1] := X_D;
aPolygon[4, 2] := Y_CD;


(************************************************************
    CREATE POLYGON STRING
*************************************************************)

sPolygonPoints := '';

FOR i := 1 TO 4 DO

    sPolygonPoints := CONCAT(
        sPolygonPoints,
        INT_TO_STRING(aPolygon[i, 1])
    );

    sPolygonPoints := CONCAT(
        sPolygonPoints,
        ','
    );

    sPolygonPoints := CONCAT(
        sPolygonPoints,
        INT_TO_STRING(aPolygon[i, 2])
    );

    IF i < 4 THEN

        sPolygonPoints := CONCAT(
            sPolygonPoints,
            ' '
        );

    END_IF;

END_FOR;

PlanarHMIWall := TRUE;
END_METHOD

METHOD WristHMIWall : BOOL
VAR
 
i : INT;
	bWristSetBlocked: BOOL := FALSE;
END_VAR

(************************************************************
    WRIST WALL BUTTON RISING EDGE DETECTION
*************************************************************)

fbRightWristWallTrig(
    CLK := GVL_HMI.RightWristWall_But
);

fbLeftWristWallTrig(
    CLK := GVL_HMI.LeftWristWall_But
);

fbWristSetTrig(
    CLK := GVL_HMI.SETWristWall_But
);

bWristSetRisingEdge := fbWristSetTrig.Q;


(************************************************************
    INITIALIZE WRIST POLYGON ONLY ONCE
*************************************************************)

IF NOT bWristPolygonInitialized THEN

    // Point A - predefined
    aWristPolygon[1, 1] := 100.0;
    aWristPolygon[1, 2] := 0.0;

    // Point B - predefined
    aWristPolygon[2, 1] := 100.0;
    aWristPolygon[2, 2] := 0.0;

    // Point C - constant
    aWristPolygon[3, 1] := 100.0;
    aWristPolygon[3, 2] := 100.0;

    bWristPolygonInitialized := TRUE;

END_IF;


(************************************************************
    SELECT WRIST WALL

    Select a new wall ONLY when no wall is active.

    WristWall:
        0 = No wall selected
        1 = Right wall selected
        2 = Left wall selected
*************************************************************)

IF WristWall = 0 THEN

    IF fbRightWristWallTrig.Q THEN

        WristWall := 1;

    ELSIF fbLeftWristWallTrig.Q THEN

        WristWall := 2;

    END_IF;

END_IF;


(************************************************************
    CONVERT ACTUAL WRIST ANGLE
    FROM DEGREES TO RADIANS
*************************************************************)

fAngleRad :=
    GVL_HMI.EndeffectorPositionPixcelUnit_Theta
    * 3.14159265359 / 180.0;


(************************************************************
    CALCULATE MOVING ENDPOINT OF PURPLE LINE

    IMPORTANT:
    This calculation runs every PLC cycle.

    The purple line follows the wrist angle
    independently of the green polygon.
*************************************************************)

fWristLineX :=
    fWristCenterX
    + fWristRadius * SIN(fAngleRad);

fWristLineY :=
    fWristCenterY
    - fWristRadius * COS(fAngleRad);


(************************************************************
    WRIST VIRTUAL WALL

    WristWall = 0:
        Keep polygon points A and B fixed.

    WristWall = 1:
        Point A follows the purple line.

    WristWall = 2:
        Point B follows the purple line.
*************************************************************)

CASE WristWall OF

    (********************************************************
        0: NO WALL ACTIVE

        Do not update polygon points A or B.

        This keeps the green area fixed after SET.
    *********************************************************)

    0:

        bWristSetEnable := FALSE;
        bWristWallInvalid := FALSE;


    (********************************************************
        1: RIGHT WALL ACTIVE

        Point A follows the purple line.
    *********************************************************)

    1:

        // Update Point A
        aWristPolygon[1, 1] := fWristLineX;
        aWristPolygon[1, 2] := fWristLineY;

        // Check wall direction
        IF aWristPolygon[1, 1] <
           aWristPolygon[2, 1] THEN

            bWristWallInvalid := FALSE;
            bWristSetEnable := TRUE;

        ELSE

            bWristWallInvalid := TRUE;
            bWristSetEnable := FALSE;

        END_IF;


    (********************************************************
        2: LEFT WALL ACTIVE

        Point B follows the purple line.
    *********************************************************)

    2:

        // Update Point B
        aWristPolygon[2, 1] := fWristLineX;
        aWristPolygon[2, 2] := fWristLineY;

        // Check wall direction
        IF aWristPolygon[1, 1] <
           aWristPolygon[2, 1] THEN

            bWristWallInvalid := FALSE;
            bWristSetEnable := TRUE;

        ELSE

            bWristWallInvalid := TRUE;
            bWristSetEnable := FALSE;

        END_IF;

END_CASE;


(************************************************************
    CHECK WHETHER SET IS BLOCKED

    TRUE means:
        - SET was pressed
        - A wall is selected
        - The selected position is invalid
*************************************************************)

bWristSetBlocked :=
    bWristSetRisingEdge
    AND (WristWall <> 0)
    AND NOT bWristSetEnable;


(************************************************************
    WHEN SET IS PRESSED, FIX THE WRIST WALL

    Similar to planar virtual wall:

    1. Keep the current polygon coordinates.
    2. Stop updating the selected boundary.
    3. Reset the wall selection.
    4. Continue updating the purple line independently.
*************************************************************)

IF bWristSetRisingEdge THEN

    IF (WristWall <> 0)
       AND bWristSetEnable THEN

        // Stop editing the current wall
        WristWall := 0;

        // Disable SET until another wall is selected
        bWristSetEnable := FALSE;

        // Clear invalid indication
        bWristWallInvalid := FALSE;

        // Deselect Right and Left buttons
        GVL_HMI.RightWristWall_But := FALSE;
        GVL_HMI.LeftWristWall_But := FALSE;

    END_IF;

    // Reset SET command
    GVL_HMI.SETWristWall_But := FALSE;

END_IF;


(************************************************************
    POINT C IS ALWAYS CONSTANT

    Point C represents the wrist rotation center.
*************************************************************)

aWristPolygon[3, 1] := fWristCenterX;
aWristPolygon[3, 2] := fWristCenterY;


(************************************************************
    CREATE POLYGON STRING FOR TWINCAT HMI

    The green polygon uses the saved coordinates
    of Points A and B.

    It does NOT directly use fWristLineX or
    fWristLineY.

    Therefore, when WristWall = 0,
    the green polygon remains fixed.
*************************************************************)

sWristPolygonPoints := '';

FOR i := 1 TO 3 DO

    // Add polygon X coordinate
    sWristPolygonPoints := CONCAT(
        sWristPolygonPoints,
        LREAL_TO_STRING(aWristPolygon[i, 1])
    );

    sWristPolygonPoints := CONCAT(
        sWristPolygonPoints,
        ','
    );

    // Add polygon Y coordinate
    sWristPolygonPoints := CONCAT(
        sWristPolygonPoints,
        LREAL_TO_STRING(aWristPolygon[i, 2])
    );

    // Add constant point after Point A
    IF i = 1 THEN

        sWristPolygonPoints := CONCAT(
            sWristPolygonPoints,
            ' 100.0,-20.0'
        );

    END_IF;

    // Add space between polygon points
    IF i < 3 THEN

        sWristPolygonPoints := CONCAT(
            sWristPolygonPoints,
            ' '
        );

    END_IF;

END_FOR;


(************************************************************
    ENABLE / UPDATE HMI POLYGON
*************************************************************)

WristHMIWall := TRUE;
END_METHOD

END_FUNCTION_BLOCK

// ---- POUs/PeelerGame/FB_PeelingGame.TcPOU
FUNCTION_BLOCK FB_PeelingGame
VAR_INPUT
	bEnable    : BOOL;
    stCartesianPosePercentage : ST_CartesianPose; // 0-100% position from Kinematics
	CartesianForcefY            : LREAL ; 
 //   RehabilitationController: E_ControllerType;
	CartesianVy : LREAL;
	
END_VAR
VAR_OUTPUT
	stJointTargetTorque : ST_JointTorque;
END_VAR
VAR
	stToUnity   : ST_PeelerToUnity;   
    stFromUnity : ST_PeelerFromUnity;
	FYThreshold    : REAL := 2.0 ;  // Minimum Force to create Resistive Force;
	VYThreshold : LREAL := 10.0;
	

END_VAR



IF bEnable THEN
    stToUnity.fY           := stCartesianPosePercentage.Y;
    stToUnity.GameIsActive := TRUE;

    // Check if close button was pressed in Unity
    IF stFromUnity.bGameFinished THEN
        stToUnity.GameIsActive := FALSE;
        stJointTargetTorque.M1 := 0.0;
        stJointTargetTorque.M2 := 0.0;
        stJointTargetTorque.M3 := 0.0;
    ELSE
        // Apply resistance ONLY when touching fruit AND moving forward (+Y)
        IF  (CartesianVy> VYThreshold )AND( CartesianForcefY > FYThreshold) THEN
            CASE stFromUnity.nObjectType OF
                1: // KIWI
                    stJointTargetTorque.M1 := 0.0;
                    stJointTargetTorque.M2 := -5.0;
                    stJointTargetTorque.M3 := 5.0;
                    
                2: // Orange
                    stJointTargetTorque.M1 := 0.0;
                    stJointTargetTorque.M2 := -10.0;
                    stJointTargetTorque.M3 := 10.0;
                    
                3: // Grapefruit
                    stJointTargetTorque.M1 := 0.0;
                    stJointTargetTorque.M2 := -15.0;
                    stJointTargetTorque.M3 := 15.0;

                4: // Melon
                    stJointTargetTorque.M1 := 0.0;
                    stJointTargetTorque.M2 := -20.0;
                    stJointTargetTorque.M3 := 20.0;

                5: // PINEAPPLE
                    stJointTargetTorque.M1 := 0.0;
                    stJointTargetTorque.M2 := -25.0;
                    stJointTargetTorque.M3 := 25.0;

                ELSE
                    stJointTargetTorque.M1 := 0.0;
                    stJointTargetTorque.M2 := 0.0;
                    stJointTargetTorque.M3 := 0.0;
            END_CASE
        ELSE
            // Zero torque if not touching, moving backwards (-Y), or stationary
            stJointTargetTorque.M1 := 0.0;
            stJointTargetTorque.M2 := 0.0;
            stJointTargetTorque.M3 := 0.0;
        END_IF
    END_IF

ELSE
    stToUnity.GameIsActive := FALSE;
    stJointTargetTorque.M1 := 0.0;
    stJointTargetTorque.M2 := 0.0;
    stJointTargetTorque.M3 := 0.0;
END_IF

END_FUNCTION_BLOCK

// ---- POUs/HardwareWallCheck.TcPOU
FUNCTION_BLOCK HardwareWallCheck
VAR_INPUT
END_VAR
VAR_OUTPUT
	HardwareActive : BOOL;
END_VAR
VAR
	SwTheta1: BOOL;
	SwTheta2: BOOL;
	SwR1: BOOL;
	SwR2: BOOL;
	SwBeta1: BOOL;
	SwBeta2: BOOL;
	
	// RTIG Function
	RtrigSwTheta1: R_TRIG;
	RtrigSwTheta2: R_TRIG;
	RtrigSwR1: R_TRIG;
	RtrigSwR2: R_TRIG;
	RtrigSwBeta1: R_TRIG;
	RtrigSwBeta2: R_TRIG;
	Activeatedswitch : ARRAY[1..6] OF BOOL;
	
END_VAR

SwTheta1 	 := (GVL_MicroSwitch.dwMicroSwitchDriverA AND 16#00020000) <> 0;  (* bit 0 *)
SwTheta2     := (GVL_MicroSwitch.dwMicroSwitchDriverA AND 16#00010000) <> 0;  (* bit 1 *)
SwR1    	 := (GVL_MicroSwitch.dwMicroSwitchDriverB AND 16#00080000) <> 0;  (* bit 0 *)
SwR2  		 := (GVL_MicroSwitch.dwMicroSwitchDriverB AND 16#00040000) <> 0;  (* bit 1 *)
SwBeta1      := (GVL_MicroSwitch.dwMicroSwitchDriverB AND 16#00020000) <> 0;  (* bit 2 *)
SwBeta2      := (GVL_MicroSwitch.dwMicroSwitchDriverB AND 16#00010000) <> 0;  (* bit 3 *)

RtrigSwBeta1(CLK :=SwBeta1);
RtrigSwBeta2(CLK :=SwBeta2);
RtrigSwR1(CLK :=SwR1);
RtrigSwR2(CLK :=SwR2);
RtrigSwTheta1(CLK :=SwTheta1);
RtrigSwTheta2(CLK :=SwTheta2);
//
Activeatedswitch[1] := RtrigSwBeta1.Q;
Activeatedswitch[2] := RtrigSwBeta2.Q;
Activeatedswitch[3] := RtrigSwR1.Q;
Activeatedswitch[4] := RtrigSwR2.Q;
Activeatedswitch[5] := RtrigSwTheta1.Q;
Activeatedswitch[6] := RtrigSwTheta2.Q;

IF (GVL_hmi.HwCheckMicroswitchLinearMax AND Activeatedswitch[3]) OR (GVL_hmi.HwCheckMicroswitchLinearMin AND Activeatedswitch[4]) OR
 (GVL_hmi.HwCheckMicroswitchRotationLeft AND Activeatedswitch[2]) OR (GVL_hmi.HwCheckMicroswitchRotationRight AND Activeatedswitch[1]) OR 
 (GVL_HMI.HwCheckMicroswitchWristLeft AND Activeatedswitch[5]) OR (GVL_HMI.HwCheckMicroswitchWristRight AND Activeatedswitch[6])

THEN

 HardwareActive := TRUE;
//ELSE
	
//	 HardwareActive := FALSE;
END_IF

END_FUNCTION_BLOCK

// ---- POUs/FB_LanguageManager.TcPOU
FUNCTION_BLOCK FB_LanguageManager
VAR_INPUT
END_VAR
VAR_OUTPUT
END_VAR
VAR
END_VAR

END_FUNCTION_BLOCK

// ---- POUs/FB_StartGame.TcPOU
FUNCTION_BLOCK FB_StartGame
VAR_INPUT
END_VAR
VAR_OUTPUT
END_VAR
VAR
END_VAR

END_FUNCTION_BLOCK

// ---- POUs/HMI_FunBlock/FB_HMI_Monitoring.TcPOU
FUNCTION_BLOCK FB_HMI_Monitoring
VAR_INPUT
END_VAR
VAR_OUTPUT
END_VAR
VAR
END_VAR

END_FUNCTION_BLOCK

// ---- GlobalTextList.TcGTLO
TEXTLIST GlobalTextList
  677 = '        rrrrtwt'
  685 = '%i'
  250 = '%s'
  652 = 'asdkfg'
  177 = 'Haji'
  25 = 'hhh'
  900 = 'salam'
  151 = 'Select Time'
  350 = 'START'
  351 = 'Status : '
END_TEXTLIST

// ---- VISUs/Screen2.TcVIS
VISUALIZATION Screen2  // 2x2
END_VISUALIZATION

// ---- VISUs/Visualization.TcVIS
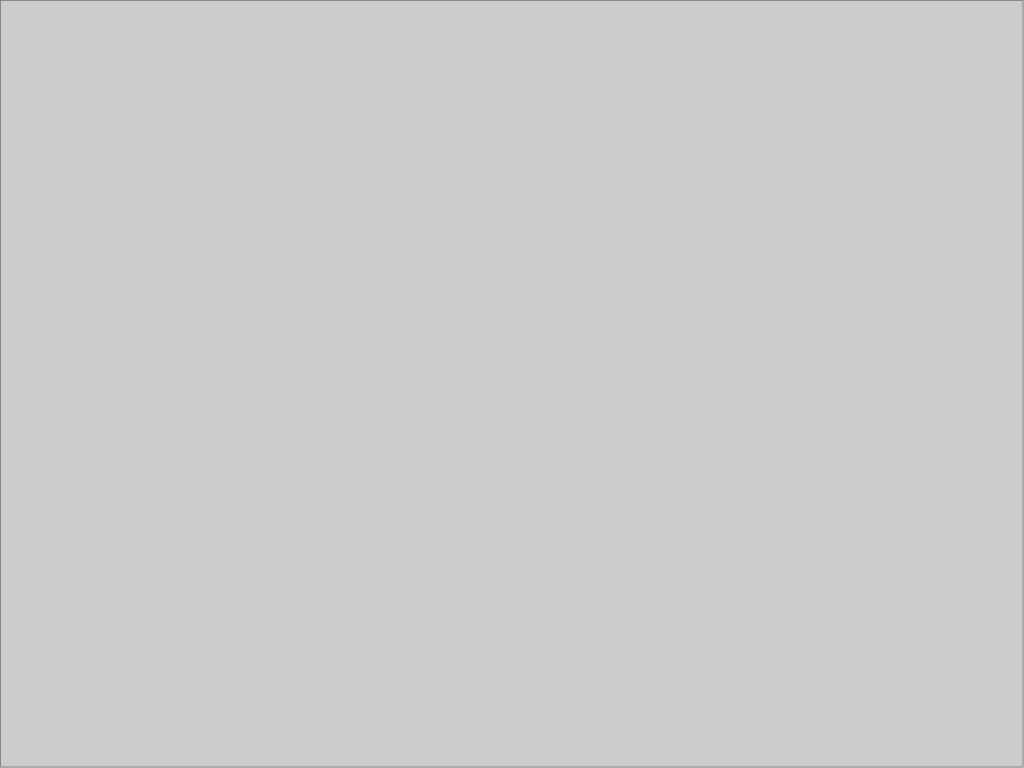
VISUALIZATION Visualization  // 1024x768
    Pie (3360,360 9280x9280)
    Pie (7150,4150 1700x1700)
    Line (8000,8440) (8000,9640)
        p3560616238: MAIN.fbKinematic.X_Visu
        p2738717112: MAIN.fbKinematic.Y_Visu
        p2858320360: MAIN.fbKinematic.Theta_Visu
    Textfield (795,6165 1100x590), "Status :"
    Textfield (775,6825 2840x430), "%s", text variable: GVL_MessageStaus.MessageStaus
    Lamp1 (3935,1815 380x410), style: Lamp-Lamp1-Yellow
END_VISUALIZATION
